(* Logix 5000 project; controller TFF vendor 1 type 14 code 107 rev 33.11; software revision 33.04; part 22 of 38 *)
(* tags used below, declared in another part *)
   Address : DINT;   // Temp Address
   Config : Configuration;   // Index Array used in configuration routines
   Index : DINT;   // Index
   TIME : DINT[2];
   AlarmAnalog : AlarmAnalog[50];   // Analog Alarm Array
   AnalogOutput : AnalogOutput[25];   // Analog Output Array
   AnalogPoint : AnalogInput[50];   // Analog Input Array
   Concentration : Concentration;
   ControlLoop : ControlLoop[20];   // Control Loop Array
   ControlLoop_FeedBagLevel : ALIAS FOR ControlLoop[2];
   ControlLoop_FeedPump : ALIAS FOR ControlLoop[1];
   ControlLoop_TIC101 : ALIAS FOR ControlLoop[7];
   Diafiltration : Diafiltration;
   DigitalPoint : DigitalPoint[150];   // Digital Point Array
   Drive : Drive[11];   // Drives Array
   FQ_Conc : ALIAS FOR Totalizer[0];   // Concentration Totalizer
   FQ_Diaf : ALIAS FOR Totalizer[1];   // DiafiltrationTotalizer
   Mixer : Mixer;   // Mixer config. structure
   Options : Options;   // Options List
   PCV101 : ALIAS FOR AnalogPoint[3];
   Phase : Phases[6];   // Phase Control Array
   Phase0_Totalizer_Feed : ALIAS FOR PhaseTotalizer[0];   // Phase 0 Total Feed
   Phase0_Totalizer_Filtrate : ALIAS FOR PhaseTotalizer[6];   // Phase 0 Total Filtrate
   Phase0_Totalizer_Transfer : ALIAS FOR PhaseTotalizer[12];   // Phase 0 Total Transfer
   Phase1_Totalizer_Feed : ALIAS FOR PhaseTotalizer[1];   // Phase 1 Total Feed
   Phase1_Totalizer_Filtrate : ALIAS FOR PhaseTotalizer[7];   // Phase 1 Total Filtrate
   Phase1_Totalizer_Transfer : ALIAS FOR PhaseTotalizer[13];   // Phase 1 Total Transfer
   Phase2_Totalizer_Feed : ALIAS FOR PhaseTotalizer[2];   // Phase 2 Total Feed
   Phase2_Totalizer_Filtrate : ALIAS FOR PhaseTotalizer[8];   // Phase 2 Total Filtrate
   Phase2_Totalizer_Transfer : ALIAS FOR PhaseTotalizer[14];   // Phase 2 Total Transfer
   Phase3_Totalizer_Feed : ALIAS FOR PhaseTotalizer[3];   // Phase 3 Total Feed
   Phase3_Totalizer_Filtrate : ALIAS FOR PhaseTotalizer[9];   // Phase 3 Total Filtrate
   Phase3_Totalizer_Transfer : ALIAS FOR PhaseTotalizer[15];   // Phase 3 Total Transfer
   Phase4_Totalizer_Feed : ALIAS FOR PhaseTotalizer[4];   // Phase 4 Total Feed
   Phase4_Totalizer_Filtrate : ALIAS FOR PhaseTotalizer[10];   // Phase 4 Total Filtrate
   Phase4_Totalizer_Transfer : ALIAS FOR PhaseTotalizer[16];   // Phase 4 Total Transfer
   Phase5_Totalizer_Feed : ALIAS FOR PhaseTotalizer[5];   // Phase 5 Total Feed
   Phase5_Totalizer_Filtrate : ALIAS FOR PhaseTotalizer[11];   // Phase 5 Total Filtrate
   Phase5_Totalizer_Transfer : ALIAS FOR PhaseTotalizer[17];   // Phase 5 Total Transfer
   Rack_Murr_Node0_Smart : IO_Station;   // Status of Node 0 Smart
   Rack_Murr_Node1_TFF : IO_Station;   // Node 1 data for MOM Config
   Rack_Murr_Node1_TFF20 : IO_Station;   // Status of Node 1 TFF20
   Rack_Murr_Node1_TFF40 : IO_Station;   // Status of Node 1 TFF40
   Rack_Murr_Node1_TFF80 : IO_Station;   // Status of Node 1 TFF80
   SIC002 : ALIAS FOR Drive[2];
   SysControl : SysControl;   // General system status and command
   Tank : TankManagement;   // Tank Management
   ThisSystem : SystemType;
   Valve : Valve[100];   // Valve Array
   ValveControl : ValveControl;   // Valve Control
   XV001 : ALIAS FOR Valve[0];
   XV002 : ALIAS FOR Valve[1];
   XV003 : ALIAS FOR Valve[2];
   XV004 : ALIAS FOR Valve[3];
   XV005 : ALIAS FOR Valve[4];
   XV006 : ALIAS FOR Valve[5];
   XV007 : ALIAS FOR Valve[6];
   XV101 : ALIAS FOR Valve[7];
   XV102 : ALIAS FOR Valve[8];
   XV201 : ALIAS FOR Valve[15];
   XV202 : ALIAS FOR Valve[16];
   XV401 : ALIAS FOR Valve[9];
   XV402 : ALIAS FOR Valve[10];
   XV403 : ALIAS FOR Valve[11];
   XV404 : ALIAS FOR Valve[12];
   XV405 : ALIAS FOR Valve[13];
   XV406 : ALIAS FOR Valve[14];
   XV701 : ALIAS FOR Valve[17];
   XV702 : ALIAS FOR Valve[18];
   XV703 : ALIAS FOR Valve[19];
   XV704 : ALIAS FOR Valve[20];
(* Process, continued *)

ROUTINE Config_IO_Station   (* structured text *)
   (* ==========================================================
   	Config I/O Station : Configure Hardware I/O Cards
   
   	Use 6 output byte for options management.
   		bit 0 to 31 : Enable / Disable 0 to 31 cards (bit index is the module number) --> 0 = Disable
   		bit 32 : Save the configuration --> 1 = Save
   		Buse Control bit 4 : 1 = Switch Off Voltage on modules , 0 = Restart the modules
   
   	List of treatments
   		- Options or configuration tools management
   		- Enable / Disable I/O modules
   		- Switch Off or restart Bus Node
   		- Module Option Management Status
   		- Module Option Management Configuration
   
   -----------------------------------------------------------------------------------------------------------------------------------------------------
   	History
   		2019-DEC-24 - Merck - Q. Spindler - Initial version for Candidate Release 1.00.00.00.a
   ============================================================*)
   
   (*Options or configuration tools management
   ============================================================*)
   
   (* Node 0 *)
   If NOT Rack_Murr_Node0_Smart.MOM_Enable_Config then
   
   	If Options.External_IO then
   		Rack_Murr_Node0_Smart.MOM_Mod_Config[3] := 0 ;
   		Rack_Murr_Node0_Smart.MOM_Mod_Config[4] := 0 ;
   		Rack_Murr_Node0_Smart.MOM_Mod_Config[5] := 0 ;
   		Rack_Murr_Node0_Smart.MOM_Mod_Config[6] := 0 ;
   	else
   		Rack_Murr_Node0_Smart.MOM_Mod_Config[3] := 1 ;
   		Rack_Murr_Node0_Smart.MOM_Mod_Config[4] := 1 ;
   		Rack_Murr_Node0_Smart.MOM_Mod_Config[5] := 1 ;
   		Rack_Murr_Node0_Smart.MOM_Mod_Config[6] := 1 ;
   	End_if ;
   
   		Rack_Murr_Node0_Smart.MOM_Mod_Config[0] := 0 ;
   		Rack_Murr_Node0_Smart.MOM_Mod_Config[1] := 0 ;
   		Rack_Murr_Node0_Smart.MOM_Mod_Config[2] := 0 ;
   		Rack_Murr_Node0_Smart.MOM_Mod_Config[7] := 0 ;
   		Rack_Murr_Node0_Smart.MOM_Mod_Config[8] := 0 ;
   		Rack_Murr_Node0_Smart.MOM_Mod_Config[9] := 0 ;
   		Rack_Murr_Node0_Smart.MOM_Mod_Config[10] := 0 ;
   		Rack_Murr_Node0_Smart.MOM_Mod_Config[11] := 0 ;
   		Rack_Murr_Node0_Smart.MOM_Mod_Config[12] := 0 ;
   		Rack_Murr_Node0_Smart.MOM_Mod_Config[13] := 0 ;
   
   	If Options.FeedTank then
   		Rack_Murr_Node0_Smart.MOM_Mod_Config[14] := 0 ;
   		Rack_Murr_Node0_Smart.MOM_Mod_Config[15] := 0 ;
   		Rack_Murr_Node0_Smart.MOM_Mod_Config[16] := 0 ;
   		Rack_Murr_Node0_Smart.MOM_Mod_Config[17] := 0 ;
   	else
   		Rack_Murr_Node0_Smart.MOM_Mod_Config[14] := 1 ;
   		Rack_Murr_Node0_Smart.MOM_Mod_Config[15] := 1 ;
   		Rack_Murr_Node0_Smart.MOM_Mod_Config[16] := 1 ;
   		Rack_Murr_Node0_Smart.MOM_Mod_Config[17] := 1 ;
   	End_if ;
   		Rack_Murr_Node0_Smart.MOM_Mod_Config[18] := 0 ;
   		Rack_Murr_Node0_Smart.MOM_Mod_Config[19] := 0 ;
   		Rack_Murr_Node0_Smart.MOM_Mod_Config[20] := 0 ;
   		Rack_Murr_Node0_Smart.MOM_Mod_Config[21] := 0 ;
   		Rack_Murr_Node0_Smart.MOM_Mod_Config[22] := 0 ;
   		Rack_Murr_Node0_Smart.MOM_Mod_Config[23] := 0 ;
   		Rack_Murr_Node0_Smart.MOM_Mod_Config[24] := 0 ;
   		Rack_Murr_Node0_Smart.MOM_Mod_Config[25] := 0 ;
   		Rack_Murr_Node0_Smart.MOM_Mod_Config[26] := 0 ;
   		Rack_Murr_Node0_Smart.MOM_Mod_Config[27] := 0 ;
   		Rack_Murr_Node0_Smart.MOM_Mod_Config[28] := 0 ;
   		Rack_Murr_Node0_Smart.MOM_Mod_Config[29] := 0 ;
   		Rack_Murr_Node0_Smart.MOM_Mod_Config[30] := 0 ;
   		Rack_Murr_Node0_Smart.MOM_Mod_Config[31] := 0 ;
   
   End_if ;
   
   
   (* Node 1 *)
   If NOT Rack_Murr_Node1_TFF.MOM_Enable_Config then
   
   	If ThisSystem.MoldType = 123 then
   		Rack_Murr_Node1_TFF.MOM_Mod_Config[0] := 0 ;
   		Rack_Murr_Node1_TFF.MOM_Mod_Config[1] := 0 ;
   		Rack_Murr_Node1_TFF.MOM_Mod_Config[2] := 0 ;
   		Rack_Murr_Node1_TFF.MOM_Mod_Config[3] := 0 ;
   		Rack_Murr_Node1_TFF.MOM_Mod_Config[4] := 0 ;
   		Rack_Murr_Node1_TFF.MOM_Mod_Config[5] := 0 ;
   		Rack_Murr_Node1_TFF.MOM_Mod_Config[6] := 0 ;
   		Rack_Murr_Node1_TFF.MOM_Mod_Config[7] := 0 ;
   		Rack_Murr_Node1_TFF.MOM_Mod_Config[8] := 0 ;
   		Rack_Murr_Node1_TFF.MOM_Mod_Config[9] := 0 ;
   		Rack_Murr_Node1_TFF.MOM_Mod_Config[10] := 0 ;
   		Rack_Murr_Node1_TFF.MOM_Mod_Config[11] := 0 ;
   		Rack_Murr_Node1_TFF.MOM_Mod_Config[12] := 0 ;
   		Rack_Murr_Node1_TFF.MOM_Mod_Config[13] := 0 ;
   		Rack_Murr_Node1_TFF.MOM_Mod_Config[14] := 0 ;
   		Rack_Murr_Node1_TFF.MOM_Mod_Config[15] := 0 ;
   		Rack_Murr_Node1_TFF.MOM_Mod_Config[16] := 0 ;
   		Rack_Murr_Node1_TFF.MOM_Mod_Config[17] := 0 ;
   		Rack_Murr_Node1_TFF.MOM_Mod_Config[18] := 0 ;
   		Rack_Murr_Node1_TFF.MOM_Mod_Config[19] := 0 ;
   		Rack_Murr_Node1_TFF.MOM_Mod_Config[20] := 0 ;
   		Rack_Murr_Node1_TFF.MOM_Mod_Config[21] := 0 ;
   		Rack_Murr_Node1_TFF.MOM_Mod_Config[22] := 0 ;
   		Rack_Murr_Node1_TFF.MOM_Mod_Config[23] := 0 ;
   		Rack_Murr_Node1_TFF.MOM_Mod_Config[24] := 0 ;
   		Rack_Murr_Node1_TFF.MOM_Mod_Config[25] := 0 ;
   		Rack_Murr_Node1_TFF.MOM_Mod_Config[26] := 0 ;
   		Rack_Murr_Node1_TFF.MOM_Mod_Config[27] := 0 ;
   		Rack_Murr_Node1_TFF.MOM_Mod_Config[28] := 0 ;
   		Rack_Murr_Node1_TFF.MOM_Mod_Config[29] := 0 ;
   		Rack_Murr_Node1_TFF.MOM_Mod_Config[30] := 0 ;
   		Rack_Murr_Node1_TFF.MOM_Mod_Config[31] := 0 ;
   	Elsif ThisSystem.MoldType = 124 then
   		Rack_Murr_Node1_TFF.MOM_Mod_Config[0] := 0 ;
   		Rack_Murr_Node1_TFF.MOM_Mod_Config[1] := 0 ;
   		Rack_Murr_Node1_TFF.MOM_Mod_Config[2] := 0 ;
   		Rack_Murr_Node1_TFF.MOM_Mod_Config[3] := 0 ;
   		Rack_Murr_Node1_TFF.MOM_Mod_Config[4] := 0 ;
   		Rack_Murr_Node1_TFF.MOM_Mod_Config[5] := 0 ;
   		Rack_Murr_Node1_TFF.MOM_Mod_Config[6] := 0 ;
   		Rack_Murr_Node1_TFF.MOM_Mod_Config[7] := 0 ;
   		Rack_Murr_Node1_TFF.MOM_Mod_Config[8] := 0 ;
   		Rack_Murr_Node1_TFF.MOM_Mod_Config[9] := 0 ;
   		Rack_Murr_Node1_TFF.MOM_Mod_Config[10] := 0 ;
   		Rack_Murr_Node1_TFF.MOM_Mod_Config[11] := 0 ;
   		Rack_Murr_Node1_TFF.MOM_Mod_Config[12] := 0 ;
   		Rack_Murr_Node1_TFF.MOM_Mod_Config[13] := 0 ;
   		Rack_Murr_Node1_TFF.MOM_Mod_Config[14] := 0 ;
   		Rack_Murr_Node1_TFF.MOM_Mod_Config[15] := 0 ;
   		Rack_Murr_Node1_TFF.MOM_Mod_Config[16] := 0 ;
   		Rack_Murr_Node1_TFF.MOM_Mod_Config[17] := 0 ;
   		Rack_Murr_Node1_TFF.MOM_Mod_Config[18] := 0 ;
   		Rack_Murr_Node1_TFF.MOM_Mod_Config[19] := 0 ;
   		Rack_Murr_Node1_TFF.MOM_Mod_Config[20] := 0 ;
   		Rack_Murr_Node1_TFF.MOM_Mod_Config[21] := 0 ;
   		Rack_Murr_Node1_TFF.MOM_Mod_Config[22] := 0 ;
   		Rack_Murr_Node1_TFF.MOM_Mod_Config[23] := 0 ;
   		Rack_Murr_Node1_TFF.MOM_Mod_Config[24] := 0 ;
   		Rack_Murr_Node1_TFF.MOM_Mod_Config[25] := 0 ;
   		Rack_Murr_Node1_TFF.MOM_Mod_Config[26] := 0 ;
   		Rack_Murr_Node1_TFF.MOM_Mod_Config[27] := 0 ;
   		Rack_Murr_Node1_TFF.MOM_Mod_Config[28] := 0 ;
   		Rack_Murr_Node1_TFF.MOM_Mod_Config[29] := 0 ;
   		Rack_Murr_Node1_TFF.MOM_Mod_Config[30] := 0 ;
   		Rack_Murr_Node1_TFF.MOM_Mod_Config[31] := 0 ;
   	Elsif ThisSystem.MoldType = 126 then
   		Rack_Murr_Node1_TFF.MOM_Mod_Config[0] := 0 ;
   		Rack_Murr_Node1_TFF.MOM_Mod_Config[1] := 0 ;
   		Rack_Murr_Node1_TFF.MOM_Mod_Config[2] := 0 ;
   		Rack_Murr_Node1_TFF.MOM_Mod_Config[3] := 0 ;
   		Rack_Murr_Node1_TFF.MOM_Mod_Config[4] := 0 ;
   		Rack_Murr_Node1_TFF.MOM_Mod_Config[5] := 0 ;
   		Rack_Murr_Node1_TFF.MOM_Mod_Config[6] := 0 ;
   		Rack_Murr_Node1_TFF.MOM_Mod_Config[7] := 0 ;
   		Rack_Murr_Node1_TFF.MOM_Mod_Config[8] := 0 ;
   		Rack_Murr_Node1_TFF.MOM_Mod_Config[9] := 0 ;
   		Rack_Murr_Node1_TFF.MOM_Mod_Config[10] := 0 ;
   		Rack_Murr_Node1_TFF.MOM_Mod_Config[11] := 0 ;
   		Rack_Murr_Node1_TFF.MOM_Mod_Config[12] := 0 ;
   		Rack_Murr_Node1_TFF.MOM_Mod_Config[13] := 0 ;
   		Rack_Murr_Node1_TFF.MOM_Mod_Config[14] := 0 ;
   		Rack_Murr_Node1_TFF.MOM_Mod_Config[15] := 0 ;
   		Rack_Murr_Node1_TFF.MOM_Mod_Config[16] := 0 ;
   		Rack_Murr_Node1_TFF.MOM_Mod_Config[17] := 0 ;
   		Rack_Murr_Node1_TFF.MOM_Mod_Config[18] := 0 ;
   		Rack_Murr_Node1_TFF.MOM_Mod_Config[19] := 0 ;
   		Rack_Murr_Node1_TFF.MOM_Mod_Config[20] := 0 ;
   		Rack_Murr_Node1_TFF.MOM_Mod_Config[21] := 0 ;
   		Rack_Murr_Node1_TFF.MOM_Mod_Config[22] := 0 ;
   		Rack_Murr_Node1_TFF.MOM_Mod_Config[23] := 0 ;
   		Rack_Murr_Node1_TFF.MOM_Mod_Config[24] := 0 ;
   		Rack_Murr_Node1_TFF.MOM_Mod_Config[25] := 0 ;
   		Rack_Murr_Node1_TFF.MOM_Mod_Config[26] := 0 ;
   		Rack_Murr_Node1_TFF.MOM_Mod_Config[27] := 0 ;
   		Rack_Murr_Node1_TFF.MOM_Mod_Config[28] := 0 ;
   		Rack_Murr_Node1_TFF.MOM_Mod_Config[29] := 0 ;
   		Rack_Murr_Node1_TFF.MOM_Mod_Config[30] := 0 ;
   		Rack_Murr_Node1_TFF.MOM_Mod_Config[31] := 0 ;
   	End_if ;
   End_if ;
   
   (*Enable / Disable I/O modules
   ============================================================*)
   
   (* Node 0 *)
   FOR Config.IndexIOMod := 0 to 7 by 1 do
   	RACK_MURR_NODE0_SMART:O.Data[0].[Config.IndexIOMod] := Rack_Murr_Node0_Smart.MOM_Mod_Config[Config.IndexIOMod] ;
   	RACK_MURR_NODE0_SMART:O.Data[1].[Config.IndexIOMod] := Rack_Murr_Node0_Smart.MOM_Mod_Config[Config.IndexIOMod+8] ;
   	RACK_MURR_NODE0_SMART:O.Data[2].[Config.IndexIOMod] := Rack_Murr_Node0_Smart.MOM_Mod_Config[Config.IndexIOMod+16] ;
   	RACK_MURR_NODE0_SMART:O.Data[3].[Config.IndexIOMod] := Rack_Murr_Node0_Smart.MOM_Mod_Config[Config.IndexIOMod+24] ;
   End_for ;
   
   (* Node 1 *)
   FOR Config.IndexIOMod := 0 to 7 by 1 do
   
   	If ThisSystem.MoldType = 123 then
   		RACK_MURR_NODE1_TFF20:O.Data[0].[Config.IndexIOMod] := Rack_Murr_Node1_TFF.MOM_Mod_Config[Config.IndexIOMod] ;
   		RACK_MURR_NODE1_TFF20:O.Data[1].[Config.IndexIOMod] := Rack_Murr_Node1_TFF.MOM_Mod_Config[Config.IndexIOMod+8] ;
   		RACK_MURR_NODE1_TFF20:O.Data[2].[Config.IndexIOMod] := Rack_Murr_Node1_TFF.MOM_Mod_Config[Config.IndexIOMod+16] ;
   		RACK_MURR_NODE1_TFF20:O.Data[3].[Config.IndexIOMod] := Rack_Murr_Node1_TFF.MOM_Mod_Config[Config.IndexIOMod+24] ;
   	Elsif ThisSystem.MoldType = 124 then
   		RACK_MURR_NODE1_TFF40:O.Data[0].[Config.IndexIOMod] := Rack_Murr_Node1_TFF.MOM_Mod_Config[Config.IndexIOMod] ;
   		RACK_MURR_NODE1_TFF40:O.Data[1].[Config.IndexIOMod] := Rack_Murr_Node1_TFF.MOM_Mod_Config[Config.IndexIOMod+8] ;
   		RACK_MURR_NODE1_TFF40:O.Data[2].[Config.IndexIOMod] := Rack_Murr_Node1_TFF.MOM_Mod_Config[Config.IndexIOMod+16] ;
   		RACK_MURR_NODE1_TFF40:O.Data[3].[Config.IndexIOMod] := Rack_Murr_Node1_TFF.MOM_Mod_Config[Config.IndexIOMod+24] ;
   	Elsif ThisSystem.MoldType = 126 then
   		RACK_MURR_NODE1_TFF80:O.Data[0].[Config.IndexIOMod] := Rack_Murr_Node1_TFF.MOM_Mod_Config[Config.IndexIOMod] ;
   		RACK_MURR_NODE1_TFF80:O.Data[1].[Config.IndexIOMod] := Rack_Murr_Node1_TFF.MOM_Mod_Config[Config.IndexIOMod+8] ;
   		RACK_MURR_NODE1_TFF80:O.Data[2].[Config.IndexIOMod] := Rack_Murr_Node1_TFF.MOM_Mod_Config[Config.IndexIOMod+16] ;
   		RACK_MURR_NODE1_TFF80:O.Data[3].[Config.IndexIOMod] := Rack_Murr_Node1_TFF.MOM_Mod_Config[Config.IndexIOMod+24] ;
   	End_if ;
   
   End_for ;
   
   (* Switch Off or restart Bus Node
   ============================================================*)
   
   (* Node 0 *)
   RACK_MURR_NODE0_SMART:O.Data[6].4 := Rack_Murr_Node0_Smart.MOM_Restart ;
   
   (* Node 1 *)
   If ThisSystem.MoldType = 123 then
   	RACK_MURR_NODE1_TFF20:O.Data[6].4 := Rack_Murr_Node1_TFF.MOM_Restart ;
   Elsif ThisSystem.MoldType = 124 then
   	RACK_MURR_NODE1_TFF40:O.Data[6].4 := Rack_Murr_Node1_TFF.MOM_Restart ;
   Elsif ThisSystem.MoldType = 126 then
   	RACK_MURR_NODE1_TFF80:O.Data[6].4 := Rack_Murr_Node1_TFF.MOM_Restart ;
   End_if ;
   
   (* Module Option Management Status
   ============================================================*)
   (* Node 0 *)
   Rack_Murr_Node0_Smart.MOM_Status := RACK_MURR_NODE0_SMART:I.Data[0];
   
   (* Node 1 *)
   If ThisSystem.MoldType = 123 then
   	Rack_Murr_Node1_TFF.MOM_Status := RACK_MURR_NODE1_TFF20:I.Data[0];
   Elsif ThisSystem.MoldType = 124 then
   	Rack_Murr_Node1_TFF.MOM_Status := RACK_MURR_NODE1_TFF40:I.Data[0];
   Elsif ThisSystem.MoldType = 126 then
   	Rack_Murr_Node1_TFF.MOM_Status := RACK_MURR_NODE1_TFF80:I.Data[0];
   End_if ;
   
   (*Module Option Management Configuration
   ============================================================*)
   
   (*save the Module Option Management configuration*)
   
   (* Node 0 *)
   RACK_MURR_NODE0_SMART:O.Data[4].0 := 1 ;
   
   (* Node 1 *)
   If ThisSystem.MoldType = 123 then
   	RACK_MURR_NODE1_TFF20:O.Data[4].0 := 1 ;
   Elsif ThisSystem.MoldType = 124 then
   	RACK_MURR_NODE1_TFF40:O.Data[4].0 := 1 ;
   Elsif ThisSystem.MoldType = 126 then
   	RACK_MURR_NODE1_TFF80:O.Data[4].0 := 1 ;
   End_if ;
   
END_ROUTINE

ROUTINE Config_Options   (* structured text *)
   (* ==========================================================
   	Config Options : Configure Options
   
   	List of treatments
   		- Configure Automatic options
   		- Configure Tank options
   		- Configure Flag for current installed clamshell
   
   -----------------------------------------------------------------------------------------------------------------------------------------------------
   	History
   		2019-DEC-24 - Merck - Q. Spindler - Initial version for Candidate Release 1.00.00.00.a
   		2022-SEP-22 - Actemium - J. Jaekel - Modification for Candidate Release 1.01.00.01.a
   				- Add Magnetic Filtrate Flowmeter instead of Ultrasonic option
   ============================================================*)
   
   (*Configure options if option Simulation mode is disabled*)
   IF Not SysControl.Simulate_Options THEN
   	// Inlet Feed Disable Option
   	IF Options.InletFeed THEN
   		Options.InletFeed_Dis := 0;
   	ELSE
   		Options.InletFeed_Dis := 1;
   	END_IF;
   
   	// No Instrum Disable Option
   	IF Options.FiltrateNoInstrum THEN
   		Options.FiltrateNoInstrum_Dis := 0;
   	ELSE
   		Options.FiltrateNoInstrum_Dis := 1;
   	END_IF;
   
   	// Tank Option
   	IF NOT Options.FeedTank THEN
   		Options.TankPH := 0;
   		Options.TankCond := 0;
   	END_IF;
   
   	// Single Use Option
   	IF Options.FiltrateNoInstrum THEN
   		Options.SingleUsePH := 0;
   	END_IF;
   
   	// Magnetic Filtrate Flowmeter instead of Ultrasonic
   	IF Options.FiltrateUltrasonicFlow THEN
   		Options.FiltrateMagneticFlow := 0;
   	ELSE
   		Options.FiltrateMagneticFlow := 1;
   	END_IF;
   END_IF;
   
   
   (*Simulate Tank Range*)
   IF Tank.Config.Simulate THEN
   
   	CASE	Tank.Config.Option_Simulate OF
   		0:	Tank.Config.Option_Current := 0 ;
   		1:	Tank.Config.Option_Current := 1 ;
   		2:	Tank.Config.Option_Current := 2 ;
   		3:	Tank.Config.Option_Current := 3 ;
   	ELSE 	Tank.Config.Option_Current := 0 ;
   	END_CASE;
   
   END_IF;
   
   (* Configure Flag for current installed clamshell
   Used to create the CCP Configuration file based on current clamshell
   ============================================================*)
   IF ThisSystem.MoldType = 123 THEN
   
   	Options.TFF20 := 1 ;
   	Options.TFF40 := 0 ;
   	Options.TFF80 := 0 ;
   
   ELSIF ThisSystem.MoldType = 124 THEN
   
   	Options.TFF20 := 0 ;
   	Options.TFF40 := 1 ;
   	Options.TFF80 := 0 ;
   
   ELSIF ThisSystem.MoldType = 126 THEN
   
   	Options.TFF20 := 0 ;
   	Options.TFF40 := 0 ;
   	Options.TFF80 := 1 ;
   
   END_IF;
END_ROUTINE

ROUTINE Config_Reset   (* structured text *)
// Set to 0  all settings
   (* ==========================================================
   	Config Reset : 	When config.reset command is activated,AnalogPoint, AlarmAnalog, AnalogOutput, Drive, DigitalPoint and Valve structure
   					are initialized to 0.
   
   	List of treatments
   		- AnalogPoint Structure reset [0] to [49]
   		- AlarmAnalog Structure reset [0] to [49]
   		- AnalogOutput Structure reset [0] to [24]
   		- Drive Structure reset [0] to [10]
   		- DigitalPoint Structure reset [0] to [149]
   		- Valve Structure reset [0] to [99]
   
   -----------------------------------------------------------------------------------------------------------------------------------------------------
   	History
   		2019-DEC-24 - Merck - Q. Spindler - Initial version for Candidate Release 1.00.00.00.a
   ============================================================*)
   
   
   (*Structure Reset [0] to [149]
   ============================================================*)
   IF Config.Reset THEN
   	FOR Config.IndexReset := 0 TO 149 BY 1 Do
   		IF Config.IndexReset <= 49 THEN
   		(*AnalogPoint Structure Reset [0] to [49]
   		====================================================*)
   			AnalogPoint[Config.IndexReset].OutofRange := 0 ;
   			AnalogPoint[Config.IndexReset].FilterType := 0 ;
   			AnalogPoint[Config.IndexReset].AveragingTotal := 0 ;
   			AnalogPoint[Config.IndexReset].Address := 0 ;
   			AnalogPoint[Config.IndexReset].RawMin := 0 ;
   			AnalogPoint[Config.IndexReset].RawMax := 0 ;
   			AnalogPoint[Config.IndexReset].RawValue := 0 ;
   			AnalogPoint[Config.IndexReset].RawLowLimit := 0 ;
   			AnalogPoint[Config.IndexReset].RawHighLimit := 0 ;
   			AnalogPoint[Config.IndexReset].FilterUser := 0 ;
   			AnalogPoint[Config.IndexReset].FilteredRaw := 0 ;
   			AnalogPoint[Config.IndexReset].FilterActual := 0 ;
   			AnalogPoint[Config.IndexReset].ScaledMin := 0 ;
   			AnalogPoint[Config.IndexReset].ScaledMax := 0 ;
   			AnalogPoint[Config.IndexReset].RangeMin := 0 ;
   			AnalogPoint[Config.IndexReset].RangeMax := 0 ;
   			AnalogPoint[Config.IndexReset].RangeMinSave := 0 ;
   			AnalogPoint[Config.IndexReset].RangeMaxSave := 0 ;
   			AnalogPoint[Config.IndexReset].RealCfg := 0 ;
   			AnalogPoint[Config.IndexReset].EnableCfg := 0 ;
   			AnalogPoint[Config.IndexReset].OverrideCfg := 0 ;
   
   		(*AlarmAnalog Structure Reset [0] to [49]
   		====================================================*)
   			AlarmAnalog[Config.IndexReset].Override := 0 ;
   			AlarmAnalog[Config.IndexReset].Disable := 0 ;
   			AlarmAnalog[Config.IndexReset].LOLODisable := 0 ;
   			AlarmAnalog[Config.IndexReset].LODisable := 0 ;
   			AlarmAnalog[Config.IndexReset].HIDisable := 0 ;
   			AlarmAnalog[Config.IndexReset].HIHIDisable := 0 ;
   			AlarmAnalog[Config.IndexReset].HIHIEnable := 0 ;
   			AlarmAnalog[Config.IndexReset].FeedPumpEnable := 0 ;
   			AlarmAnalog[Config.IndexReset].FeedPumpTag := 0 ;
   			AlarmAnalog[Config.IndexReset].TransferPumpEnable := 0 ;
   			AlarmAnalog[Config.IndexReset].TransferPumpTag := 0 ;
   			AlarmAnalog[Config.IndexReset].LOLO := 0 ;
   			AlarmAnalog[Config.IndexReset].LO := 0 ;
   			AlarmAnalog[Config.IndexReset].HI := 0 ;
   			AlarmAnalog[Config.IndexReset].HIHI := 0 ;
   			AlarmAnalog[Config.IndexReset].LOLOTimer.PRE := 0 ;
   			AlarmAnalog[Config.IndexReset].LOTimer.PRE := 0 ;
   			AlarmAnalog[Config.IndexReset].HITimer.PRE := 0 ;
   			AlarmAnalog[Config.IndexReset].HIHITimer.PRE := 0 ;
   			AlarmAnalog[Config.IndexReset].EnableCfg := 0 ;
   		End_IF;
   
   		(*AnalogOutput Structure Reset [0] to [24]
   		====================================================*)
   		IF Config.IndexReset <= 24 THEN
   			AnalogOutput[Config.IndexReset].RawValue := 0 ;
   			AnalogOutput[Config.IndexReset].RawMin := 0 ;
   			AnalogOutput[Config.IndexReset].RawMax := 0 ;
   			AnalogOutput[Config.IndexReset].ScaledMin := 0 ;
   			AnalogOutput[Config.IndexReset].ScaledMax := 0 ;
   			AnalogOutput[Config.IndexReset].EnableCfg := 0 ;
   		End_IF;
   
   		(*Drive Structure Reset [0] to [10]
   		====================================================*)
   		IF Config.IndexReset <= 10 THEN
   			Drive[Config.IndexReset].OutputAddress := 0 ;
   			Drive[Config.IndexReset].InputAddress := 0 ;
   			Drive[Config.IndexReset].RunInput := 0 ;
   			Drive[Config.IndexReset].InterlockTimer.PRE := 0 ;
   			Drive[Config.IndexReset].EnableCfg := 0 ;
   			Drive[Config.IndexReset].ReverseCfg := 0 ;
   			Drive[Config.IndexReset].Direction := 0 ;
   			Drive[Config.IndexReset].DirectionAddress := 0 ;
   		End_IF;
   
   		IF Config.IndexReset <= 99 THEN
   				(*Valves Structure Reset [0] to [99]
   		====================================================*)
   		Valve[Config.IndexReset].ZSOpenEnable := 0 ;
   		Valve[Config.IndexReset].ZSCloseEnable := 0 ;
   		Valve[Config.IndexReset].ZSOverride := 0 ;
   		Valve[Config.IndexReset].FailState := 0 ;
   		Valve[Config.IndexReset].Ports := 0 ;
   		Valve[Config.IndexReset].EnableCfg := 0 ;
   		Valve[Config.IndexReset].StatusWord := 0 ;
   		Valve[Config.IndexReset].ZSOpenAddress := 0 ;
   		Valve[Config.IndexReset].ZSCloseAddress := 0 ;
   		Valve[Config.IndexReset].OutputAddress := 0 ;
   		Valve[Config.IndexReset].AlarmTimer.PRE := 0 ;
   		Valve[Config.IndexReset].AutoCloseTimer.PRE := 0 ;
   		End_IF;
   
   		(*DigitalPoint Structure Reset [0] to [149]
   		====================================================*)
   		DigitalPoint[Config.IndexReset].Override := 0 ;
   		DigitalPoint[Config.IndexReset].DelayTimer.PRE := 0 ;
   		DigitalPoint[Config.IndexReset].Priority := 0 ;
   		DigitalPoint[Config.IndexReset].EnableCfg := 0 ;
   		DigitalPoint[Config.IndexReset].ActiveStateCFg := 0 ;
   		DigitalPoint[Config.IndexReset].RealInputCfg := 0 ;
   		DigitalPoint[Config.IndexReset].InputAddressCfg := 0 ;
   		DigitalPoint[Config.IndexReset].AlarmCfg := 0 ;
   		DigitalPoint[Config.IndexReset].AlarmStateCfg := 0 ;
   		DigitalPoint[Config.IndexReset].OverrideCfg := 0 ;
   		DigitalPoint[Config.IndexReset].PriorityCfg := 0 ;
   		DigitalPoint[Config.IndexReset].Cond1Cfg := 0 ;
   		DigitalPoint[Config.IndexReset].Cond2Cfg := 0 ;
   		DigitalPoint[Config.IndexReset].FlashingInputCfg := 0 ;
   
   	END_FOR;
   End_IF;
   (*Reset config.reset to execute routine one time*)
   Config.Reset := 0;
END_ROUTINE

ROUTINE Config_Totalizers   (* structured text *)
   (* ==========================================================
   	Config Totalizers : Configure Totalizers Structure
   
   	List of treatments
   		- Phase 0 Totalizers
   		- Phase 1 Totalizers
   		- Phase 2 Totalizers
   		- Phase 3 Totalizers
   		- Phase 4 Totalizers
   		- Phase 5 Totalizers
   		- Concentration and Diafiltration Totalizers
   
   -----------------------------------------------------------------------------------------------------------------------------------------------------
   	History
   		2019-DEC-24 - Merck - Q. Spindler - Initial version for Candidate Release 1.00.00.00.a
   		2022-JAN-11 - Merck - Q. Spindler - Modifications for Candidate Release 1.01.00.00.a
   					- Add transfer totalizers
   ============================================================*)
   
   
   (*Phase 0 Totalizers
   ============================================================*)
   Phase0_Totalizer_Feed.EnableCfg := 1 ;
   Phase0_Totalizer_Feed.SourceAddressCfg := 42 ;
   Phase0_Totalizer_Feed.SourceTypeCfg := 0 ;
   Phase0_Totalizer_Feed.PVscale := 60 ;
   
   Phase0_Totalizer_Filtrate.EnableCfg := 1 ;
   Phase0_Totalizer_Filtrate.SourceAddressCfg := 2 ;
   Phase0_Totalizer_Filtrate.SourceTypeCfg := 0 ;
   Phase0_Totalizer_Filtrate.PVscale := 60 ;
   
   Phase0_Totalizer_Transfer.EnableCfg := 1 ;
   Phase0_Totalizer_Transfer.SourceAddressCfg := 20 ;
   Phase0_Totalizer_Transfer.SourceTypeCfg := 0 ;
   Phase0_Totalizer_Transfer.PVscale := 60 ;
   
   (*Phase 1 Totalizers
   ============================================================*)
   Phase1_Totalizer_Feed.EnableCfg := 1 ;
   Phase1_Totalizer_Feed.SourceAddressCfg := 42 ;
   Phase1_Totalizer_Feed.SourceTypeCfg := 0 ;
   Phase1_Totalizer_Feed.PVscale := 60 ;
   
   Phase1_Totalizer_Filtrate.EnableCfg := 1 ;
   Phase1_Totalizer_Filtrate.SourceAddressCfg := 2 ;
   Phase1_Totalizer_Filtrate.SourceTypeCfg := 0 ;
   Phase1_Totalizer_Filtrate.PVscale := 60 ;
   
   Phase1_Totalizer_Transfer.EnableCfg := 1 ;
   Phase1_Totalizer_Transfer.SourceAddressCfg := 20 ;
   Phase1_Totalizer_Transfer.SourceTypeCfg := 0 ;
   Phase1_Totalizer_Transfer.PVscale := 60 ;
   
   (*Phase 2 Totalizers
   ============================================================*)
   Phase2_Totalizer_Feed.EnableCfg := 1 ;
   Phase2_Totalizer_Feed.SourceAddressCfg := 42 ;
   Phase2_Totalizer_Feed.SourceTypeCfg := 0 ;
   Phase2_Totalizer_Feed.PVscale := 60 ;
   
   Phase2_Totalizer_Filtrate.EnableCfg := 1 ;
   Phase2_Totalizer_Filtrate.SourceAddressCfg := 2 ;
   Phase2_Totalizer_Filtrate.SourceTypeCfg := 0 ;
   Phase2_Totalizer_Filtrate.PVscale := 60 ;
   
   Phase2_Totalizer_Transfer.EnableCfg := 1 ;
   Phase2_Totalizer_Transfer.SourceAddressCfg := 20 ;
   Phase2_Totalizer_Transfer.SourceTypeCfg := 0 ;
   Phase2_Totalizer_Transfer.PVscale := 60 ;
   
   (*Phase 3 Totalizers
   ============================================================*)
   Phase3_Totalizer_Feed.EnableCfg := 1 ;
   Phase3_Totalizer_Feed.SourceAddressCfg := 42 ;
   Phase3_Totalizer_Feed.SourceTypeCfg := 0 ;
   Phase3_Totalizer_Feed.PVscale := 60 ;
   
   Phase3_Totalizer_Filtrate.EnableCfg := 1 ;
   Phase3_Totalizer_Filtrate.SourceAddressCfg := 2 ;
   Phase3_Totalizer_Filtrate.SourceTypeCfg := 0 ;
   Phase3_Totalizer_Filtrate.PVscale := 60 ;
   
   Phase3_Totalizer_Transfer.EnableCfg := 1 ;
   Phase3_Totalizer_Transfer.SourceAddressCfg := 20 ;
   Phase3_Totalizer_Transfer.SourceTypeCfg := 0 ;
   Phase3_Totalizer_Transfer.PVscale := 60 ;
   
   (*Phase 4 Totalizers
   ============================================================*)
   Phase4_Totalizer_Feed.EnableCfg := 1 ;
   Phase4_Totalizer_Feed.SourceAddressCfg := 42 ;
   Phase4_Totalizer_Feed.SourceTypeCfg := 0 ;
   Phase4_Totalizer_Feed.PVscale := 60 ;
   
   Phase4_Totalizer_Filtrate.EnableCfg := 1 ;
   Phase4_Totalizer_Filtrate.SourceAddressCfg := 2 ;
   Phase4_Totalizer_Filtrate.SourceTypeCfg := 0 ;
   Phase4_Totalizer_Filtrate.PVscale := 60 ;
   
   Phase4_Totalizer_Transfer.EnableCfg := 1 ;
   Phase4_Totalizer_Transfer.SourceAddressCfg := 20 ;
   Phase4_Totalizer_Transfer.SourceTypeCfg := 0 ;
   Phase4_Totalizer_Transfer.PVscale := 60 ;
   
   (*Phase 5 Totalizers
   ============================================================*)
   Phase5_Totalizer_Feed.EnableCfg := 1 ;
   Phase5_Totalizer_Feed.SourceAddressCfg := 42 ;
   Phase5_Totalizer_Feed.SourceTypeCfg := 0 ;
   Phase5_Totalizer_Feed.PVscale := 60 ;
   
   Phase5_Totalizer_Filtrate.EnableCfg := 1 ;
   Phase5_Totalizer_Filtrate.SourceAddressCfg := 2 ;
   Phase5_Totalizer_Filtrate.SourceTypeCfg := 0 ;
   Phase5_Totalizer_Filtrate.PVscale := 60 ;
   
   Phase5_Totalizer_Transfer.EnableCfg := 1 ;
   Phase5_Totalizer_Transfer.SourceAddressCfg := 20 ;
   Phase5_Totalizer_Transfer.SourceTypeCfg := 0 ;
   Phase5_Totalizer_Transfer.PVscale := 60 ;
   
   (*Concentration and Diafiltration Totalizers
   ============================================================*)
   
   FQ_Conc.PVscale := 60 ;
   FQ_Diaf.PVscale := 60 ;
END_ROUTINE

ROUTINE Config_Valve   (* structured text *)
// Apply the default configuration
   (* ==========================================================
   	Config Valve : Configure Valve Structure
   
   	List of treatments
   		- Valve[0] : Valve XV001
   		- Valve[1] : Valve XV002
   		- Valve[2] : Valve XV003
   		- Valve[3] : Valve XV004
   		- Valve[4] : Valve XV005
   		- Valve[5] : Valve XV006
   		- Valve[6] : Valve XV007
   		- Valve[7] : Valve XV101
   		- Valve[8] : Valve XV102
   		- Valve[9] : Valve XV401
   		- Valve[10]: Valve XV402
   		- Valve[11]: Valve XV403
   		- Valve[12]: Valve XV404
   		- Valve[13]: Valve XV405
   		- Valve[14]: Valve XV406
   		- Valve[15]: Valve XV201
   		- Valve[16]: Valve XV202
   		- Valve[17]: Valve XV701
   		- Valve[18]: Valve XV702
   		- Valve[19]: Valve XV703
   		- Valve[20]: Valve XV704
   		- Reset Loop : Set to 0 the Valve[21 to 99].EnableCfg
   
   -----------------------------------------------------------------------------------------------------------------------------------------------------
   	History
   		2019-DEC-24 - Merck - Q. Spindler - Initial version for Candidate Release 1.00.00.00.a
   		2020-APR-06 - Merck - Q. Spindler - Modifications for Candidate Release 1.00.00.00.b
   					- Invert FailState for XV201
   					- Add ZSClose for XV003,XV004,XV005,XV006,XV007
   		2020-JUN-19 - Merck - Q. Spindler - Modifications for Candidate Release 1.00.00.00.c
   					- Change ZSClose to ZSOpen for XV003,XV004,XV005,XV006,XV007
   ============================================================*)
   
   
   (*Max valve number use as terminal value in loop
   ============================================================*)
   ValveControl.MaxValveNum := 32;
   
   (*Valve[0] : Valve XV001
   ============================================================*)
   Valve[0].EnableCfg := 1 ;
   Valve[0].FailState := 1 ;
   Valve[0].ZSOverride := 1 ;
   Valve[0].Ports := 0 ;
   Valve[0].PriorityCfg := 0 ;
   Valve[0].ZSOpenEnable := 0 ;
   Valve[0].Alarm := 0 ;
   Valve[0].ZSCloseEnable := 0 ;
   Valve[0].ZSOpenAddress := 0 ;
   Valve[0].ZSCloseAddress := 0 ;
   Valve[0].OutputAddress := 32 ;
   
   (*Valve[1] : Valve XV002
   ============================================================*)
   Valve[1].EnableCfg := 1 ;
   Valve[1].FailState := 1 ;
   Valve[1].ZSOverride := 1 ;
   Valve[1].Ports := 0 ;
   Valve[1].PriorityCfg := 0 ;
   Valve[1].ZSOpenEnable := 0 ;
   Valve[1].Alarm := 0 ;
   Valve[1].ZSCloseEnable := 0 ;
   Valve[1].ZSOpenAddress := 0 ;
   Valve[1].ZSCloseAddress := 0 ;
   Valve[1].OutputAddress := 33 ;
   
   (*Valve[2] : Valve XV003
   ============================================================*)
   IF Options.InletFeed THEN
   	Valve[2].EnableCfg := 1 ;
   ELSE
   	Valve[2].EnableCfg := 0 ;
   	Valve[2].Alarm := 0 ;
   END_IF;
   Valve[2].FailState := 0 ;
   Valve[2].Ports := 0 ;
   Valve[2].PriorityCfg := 1 ;
   Valve[2].ZSOpenEnable := 1 ;
   Valve[2].ZSCloseEnable := 0 ;
   Valve[2].ZSOpenAddress := 2 ;
   Valve[2].ZSCloseAddress := 0 ;
   Valve[2].OutputAddress := 34 ;
   
   (*Valve[3] : Valve XV004
   ============================================================*)
   IF Options.InletFeed THEN
   	Valve[3].EnableCfg := 1 ;
   ELSE
   	Valve[3].EnableCfg := 0 ;
   	Valve[3].Alarm := 0 ;
   END_IF;
   Valve[3].FailState := 0 ;
   Valve[3].Ports := 0 ;
   Valve[3].PriorityCfg := 1 ;
   Valve[3].ZSOpenEnable := 1 ;
   Valve[3].ZSCloseEnable := 0 ;
   Valve[3].ZSOpenAddress := 3 ;
   Valve[3].ZSCloseAddress := 0 ;
   Valve[3].OutputAddress := 35 ;
   
   (*Valve[4] : Valve XV005
   ============================================================*)
   IF Options.InletFeed THEN
   	Valve[4].EnableCfg := 1 ;
   ELSE
   	Valve[4].EnableCfg := 0 ;
   	Valve[4].Alarm := 0 ;
   END_IF;
   Valve[4].FailState := 0 ;
   Valve[4].Ports := 0 ;
   Valve[4].PriorityCfg := 1 ;
   Valve[4].ZSOpenEnable := 1 ;
   Valve[4].ZSCloseEnable := 0 ;
   Valve[4].ZSOpenAddress := 4 ;
   Valve[4].ZSCloseAddress := 0 ;
   Valve[4].OutputAddress := 36 ;
   
   (*Valve[5] : Valve XV006
   ============================================================*)
   IF Options.InletFeed THEN
   	Valve[5].EnableCfg := 1 ;
   ELSE
   	Valve[5].EnableCfg := 0 ;
   	Valve[5].Alarm := 0 ;
   END_IF;
   Valve[5].FailState := 0 ;
   Valve[5].Ports := 0 ;
   Valve[5].PriorityCfg := 1 ;
   Valve[5].ZSOpenEnable := 1 ;
   Valve[5].ZSCloseEnable := 0 ;
   Valve[5].ZSOpenAddress := 5 ;
   Valve[5].ZSCloseAddress := 0 ;
   Valve[5].OutputAddress := 37 ;
   
   (*Valve[6] : Valve XV007
   ============================================================*)
   IF Options.InletFeed THEN
   	Valve[6].EnableCfg := 1 ;
   ELSE
   	Valve[6].EnableCfg := 0 ;
   	Valve[6].Alarm := 0 ;
   END_IF;
   Valve[6].FailState := 0 ;
   Valve[6].Ports := 0 ;
   Valve[6].PriorityCfg := 1 ;
   Valve[6].ZSOpenEnable := 1 ;
   Valve[6].ZSCloseEnable := 0 ;
   Valve[6].ZSOpenAddress := 6;
   Valve[6].ZSCloseAddress := 0 ;
   Valve[6].OutputAddress := 38 ;
   
   (*Valve[7] : Valve XV101
   ============================================================*)
   Valve[7].EnableCfg := 1 ;
   Valve[7].FailState := 1 ;
   Valve[7].ZSOverride := 1 ;
   Valve[7].Ports := 0 ;
   Valve[7].PriorityCfg := 0 ;
   Valve[7].ZSOpenEnable := 0 ;
   Valve[7].Alarm := 0 ;
   Valve[7].ZSCloseEnable := 0 ;
   Valve[7].ZSOpenAddress := 0 ;
   Valve[7].ZSCloseAddress := 0 ;
   Valve[7].OutputAddress := 39 ;
   
   (*Valve[8] : Valve XV102
   ============================================================*)
   Valve[8].EnableCfg := 1 ;
   Valve[8].FailState := 1 ;
   Valve[8].ZSOverride := 1 ;
   Valve[8].Ports := 0 ;
   Valve[8].PriorityCfg := 0 ;
   Valve[8].ZSOpenEnable := 0 ;
   Valve[8].Alarm := 0 ;
   Valve[8].ZSCloseEnable := 0 ;
   Valve[8].ZSOpenAddress := 0 ;
   Valve[8].ZSCloseAddress := 0 ;
   Valve[8].OutputAddress := 40 ;
   
   (*Valve[9] : Valve XV401
   ============================================================*)
   Valve[9].EnableCfg := 1 ;
   Valve[9].FailState := 0 ;
   Valve[9].ZSOverride := 1 ;
   Valve[9].Ports := 0 ;
   Valve[9].PriorityCfg := 0 ;
   Valve[9].ZSOpenEnable := 0 ;
   Valve[9].Alarm := 0 ;
   Valve[9].ZSCloseEnable := 0 ;
   Valve[9].ZSOpenAddress := 0 ;
   Valve[9].ZSCloseAddress := 0 ;
   Valve[9].OutputAddress := 41 ;
   
   (*Valve[10]: Valve XV402
   ============================================================*)
   Valve[10].EnableCfg := 1 ;
   Valve[10].FailState := 0 ;
   Valve[10].ZSOverride := 1 ;
   Valve[10].Ports := 0 ;
   Valve[10].PriorityCfg := 0 ;
   Valve[10].ZSOpenEnable := 0 ;
   Valve[10].Alarm := 0 ;
   Valve[10].ZSCloseEnable := 0 ;
   Valve[10].ZSOpenAddress := 0 ;
   Valve[10].ZSCloseAddress := 0 ;
   Valve[10].OutputAddress := 42 ;
   
   (*Valve[11]: Valve XV403
   ============================================================*)
   Valve[11].EnableCfg := 1 ;
   Valve[11].FailState := 0 ;
   Valve[11].ZSOverride := 1 ;
   Valve[11].Ports := 0 ;
   Valve[11].PriorityCfg := 0 ;
   Valve[11].ZSOpenEnable := 0 ;
   Valve[11].Alarm := 0 ;
   Valve[11].ZSCloseEnable := 0 ;
   Valve[11].ZSOpenAddress := 0 ;
   Valve[11].ZSCloseAddress := 0 ;
   Valve[11].OutputAddress := 43 ;
   
   (*Valve[12]: Valve XV404
   ============================================================*)
   Valve[12].EnableCfg := 1 ;
   Valve[12].FailState := 0 ;
   Valve[12].ZSOverride := 1 ;
   Valve[12].Ports := 0 ;
   Valve[12].PriorityCfg := 0 ;
   Valve[12].ZSOpenEnable := 0 ;
   Valve[12].Alarm := 0 ;
   Valve[12].ZSCloseEnable := 0 ;
   Valve[12].ZSOpenAddress := 0 ;
   Valve[12].ZSCloseAddress := 0 ;
   Valve[12].OutputAddress := 44 ;
   
   (*Valve[13]: Valve XV405
   ============================================================*)
   IF Options.InletFeed THEN
   	Valve[13].EnableCfg := 0 ;
   ELSE
   	Valve[13].EnableCfg := 1 ;
   END_IF;
   Valve[13].FailState := 0 ;
   Valve[13].ZSOverride := 1 ;
   Valve[13].Ports := 0 ;
   Valve[13].PriorityCfg := 0 ;
   Valve[13].ZSOpenEnable := 0 ;
   Valve[13].Alarm := 0 ;
   Valve[13].ZSCloseEnable := 0 ;
   Valve[13].ZSOpenAddress := 0 ;
   Valve[13].ZSCloseAddress := 0 ;
   Valve[13].OutputAddress := 45 ;
   
   (*Valve[14]: Valve XV406
   ============================================================*)
   IF Options.InletFeed THEN
   	Valve[14].EnableCfg := 0 ;
   ELSE
   	Valve[14].EnableCfg := 1 ;
   END_IF;
   Valve[14].FailState := 0 ;
   Valve[14].ZSOverride := 1 ;
   Valve[14].Ports := 0 ;
   Valve[14].PriorityCfg := 0 ;
   Valve[14].ZSOpenEnable := 0 ;
   Valve[14].Alarm := 0 ;
   Valve[14].ZSCloseEnable := 0 ;
   Valve[14].ZSOpenAddress := 0 ;
   Valve[14].ZSCloseAddress := 0 ;
   Valve[14].OutputAddress := 46 ;
   
   (*Valve[15]: Valve XV201
   ============================================================*)
   Valve[15].EnableCfg := 1 ;
   Valve[15].FailState := 0 ;
   Valve[15].ZSOverride := 1 ;
   Valve[15].Ports := 0 ;
   Valve[15].PriorityCfg := 0 ;
   Valve[15].ZSOpenEnable := 0 ;
   Valve[15].Alarm := 0 ;
   Valve[15].ZSCloseEnable := 0 ;
   Valve[15].ZSOpenAddress := 0 ;
   Valve[15].ZSCloseAddress := 0 ;
   Valve[15].OutputAddress := 47 ;
   
   (*Valve[16]: Valve XV202
   ============================================================*)
   Valve[16].EnableCfg := 1 ;
   Valve[16].FailState := 0 ;
   Valve[16].ZSOverride := 1 ;
   Valve[16].Ports := 0 ;
   Valve[16].PriorityCfg := 0 ;
   Valve[16].ZSOpenEnable := 0 ;
   Valve[16].Alarm := 0 ;
   Valve[16].ZSCloseEnable := 0 ;
   Valve[16].ZSOpenAddress := 0 ;
   Valve[16].ZSCloseAddress := 0 ;
   Valve[16].OutputAddress := 48 ;
   
   (*Valve[17]: Valve XV701
   ============================================================*)
   Valve[17].EnableCfg := 1 ;
   Valve[17].FailState := 0 ;
   Valve[17].ZSOverride := 1 ;
   Valve[17].Ports := 0 ;
   Valve[17].PriorityCfg := 0 ;
   Valve[17].ZSOpenEnable := 0 ;
   Valve[17].Alarm := 0 ;
   Valve[17].ZSCloseEnable := 0 ;
   Valve[17].ZSOpenAddress := 0 ;
   Valve[17].ZSCloseAddress := 0 ;
   Valve[17].OutputAddress := 49 ;
   
   (*Valve[18]: Valve XV702
   ============================================================*)
   Valve[18].EnableCfg := 1 ;
   Valve[18].FailState := 0 ;
   Valve[18].ZSOverride := 1 ;
   Valve[18].Ports := 0 ;
   Valve[18].PriorityCfg := 0 ;
   Valve[18].ZSOpenEnable := 0 ;
   Valve[18].Alarm := 0 ;
   Valve[18].ZSCloseEnable := 0 ;
   Valve[18].ZSOpenAddress := 0 ;
   Valve[18].ZSCloseAddress := 0 ;
   Valve[18].OutputAddress := 50 ;
   
   (*Valve[19]: Valve XV703
   ============================================================*)
   Valve[19].EnableCfg := 1 ;
   Valve[19].FailState := 0 ;
   Valve[19].ZSOverride := 1 ;
   Valve[19].Ports := 0 ;
   Valve[19].PriorityCfg := 0 ;
   Valve[19].ZSOpenEnable := 0 ;
   Valve[19].Alarm := 0 ;
   Valve[19].ZSCloseEnable := 0 ;
   Valve[19].ZSOpenAddress := 0 ;
   Valve[19].ZSCloseAddress := 0 ;
   Valve[19].OutputAddress := 51 ;
   
   (*Valve[20]: Valve XV704
   ============================================================*)
   Valve[20].EnableCfg := 1 ;
   Valve[20].FailState := 0 ;
   Valve[20].ZSOverride := 1 ;
   Valve[20].Ports := 0 ;
   Valve[20].PriorityCfg := 0 ;
   Valve[20].ZSOpenEnable := 0 ;
   Valve[20].Alarm := 0 ;
   Valve[20].ZSCloseEnable := 0 ;
   Valve[20].ZSOpenAddress := 0 ;
   Valve[20].ZSCloseAddress := 0 ;
   Valve[20].OutputAddress := 52 ;
   
   (*Reset Loop : Set to 0 the Valve[21 to 99].EnableCfg
   ============================================================*)
   FOR Config.IndeXValve := 21 to 99 by 1 do
   	Valve[Config.IndeXValve].EnableCfg := 0 ;
   	Valve[Config.IndeXValve].Alarm := 0 ;
   	Valve[Config.IndeXValve].Control := 0 ;
   	Valve[Config.IndeXValve].Auto := 0 ;
   	Valve[Config.IndeXValve].Manual := 0 ;
   	Valve[Config.IndeXValve].StatusWord := 0 ;
   	Valve[Config.IndeXValve].Status := 0 ;
   End_for ;
END_ROUTINE

ROUTINE Control_Loop   (* ladder *)
// Control Loop Routine
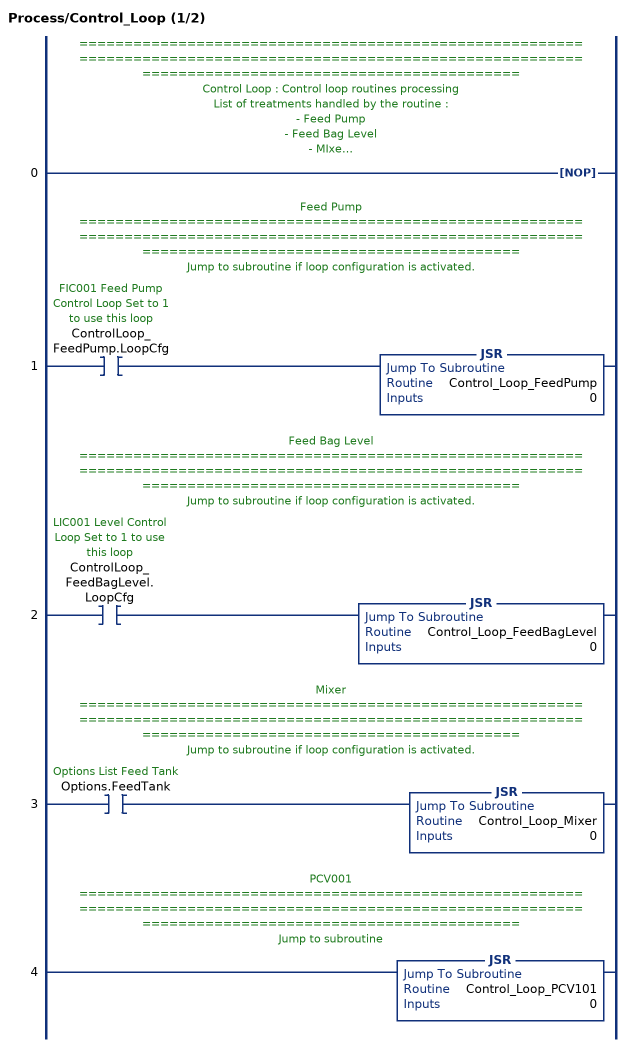
   // ==========================================================================================================================================================
   //                                                                                                                 Control Loop : Control loop routines processing
   //                                                     List of treatments handled by the routine :
   //                                                          - Feed Pump
   //                                                          - Feed Bag Level
   //                                                          - MIxer
   //                                                          - PCV001
   //                                                           - PCV101
   //                                                          - TIC101
   //                                                     -----------------------------------------------------------------------------------------------------------------------------------------------------
   //                                                     History
   // 		2019-DEC-24 - Merck - Q. Spindler - Initial version for Candidate Release 1.00.00.00.a
   // ==========================================================================================================================================================
   0: NOP();
   // Feed Pump
   // ==========================================================================================================================================================
   // Jump to subroutine if loop configuration is activated.
   1: XIC(ControlLoop_FeedPump.LoopCfg)JSR(Control_Loop_FeedPump,0);
   // Feed Bag Level
   // ==========================================================================================================================================================
   // Jump to subroutine if loop configuration is activated.
   2: XIC(ControlLoop_FeedBagLevel.LoopCfg)JSR(Control_Loop_FeedBagLevel,0);
   // Mixer
   // ==========================================================================================================================================================
   // Jump to subroutine if loop configuration is activated.
   3: XIC(Options.FeedTank)JSR(Control_Loop_Mixer,0);
   // PCV001
   // ==========================================================================================================================================================
   // Jump to subroutine
   4: JSR(Control_Loop_PCV101,0);
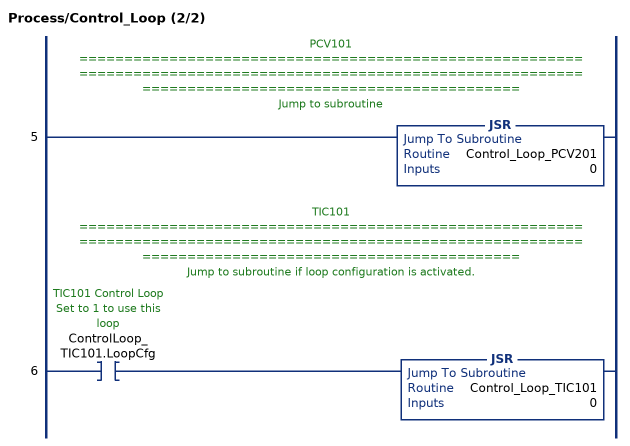
   // PCV101
   // ==========================================================================================================================================================
   // Jump to subroutine
   5: JSR(Control_Loop_PCV201,0);
   // TIC101
   // ==========================================================================================================================================================
   // Jump to subroutine if loop configuration is activated.
   6: XIC(ControlLoop_TIC101.LoopCfg)JSR(Control_Loop_TIC101,0);
END_ROUTINE

ROUTINE Control_Loop_FeedBagLevel   (* ladder *)
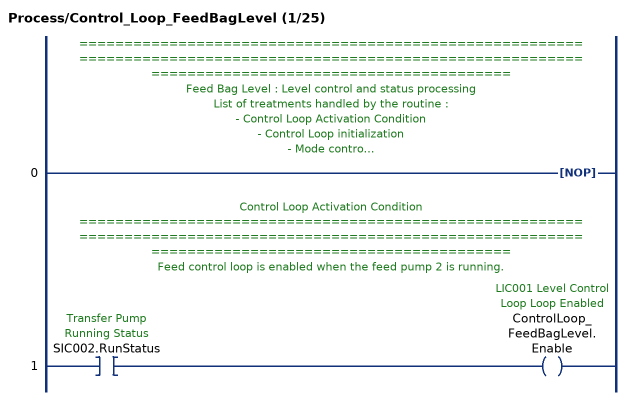
   // ========================================================================================================================================================
   //                                                                                                       Feed Bag Level : Level control and status processing
   //                                                     List of treatments handled by the routine :
   //                                                          - Control Loop Activation Condition
   //                                                          - Control Loop initialization
   //                                                          - Mode control
   //                                                          - Control Loop deadband calculation
   //                                                          - Management of ramping control
   //                                                          - Control Loop Stability control
   //                                                          - Control Loop manual state control
   //                                                          - Management of PID instruction
   //                                                          - Control of the analog output
   //                                                     -----------------------------------------------------------------------------------------------------------------------------------------------------
   //                                                     History
   //                		2019-DEC-24 - Merck - Q. Spindler - Initial version for Candidate Release 1.00.00.00.a
   // 		2020-SEP-09 - Merck - Q. Spindler - Modifications for Candidate Release 1.00.00.00.d
   // 					- Add ControlLoop Enable and not manual condition for DBOK status
   //                    - Set ramp rate minimum to 0.1
   // 		2021-APR-16 - Merck - Q. Spindler - Modifications for Candidate Release 1.00.00.00.e
   //                                        - Add Initialize address if no mode selected.
   //                                                              - The wrong control loop was used in the PID initialisation
   // 		2022-NOV-21 - Actemium - J. Jaekel - Modifications for Candidate Release 1.01.00.01.b
   // - Set manuel mode if Auto Mode 2 is enabled and TransferFlow option is disabled.
   // - If no mode is active, activate the manual mode.
   // ========================================================================================================================================================
   0: NOP();
   // Control Loop Activation Condition
   // ========================================================================================================================================================
   // Feed control loop is enabled when the feed pump 2 is running.
   1: XIC(SIC002.RunStatus)OTE(ControlLoop_FeedBagLevel.Enable);
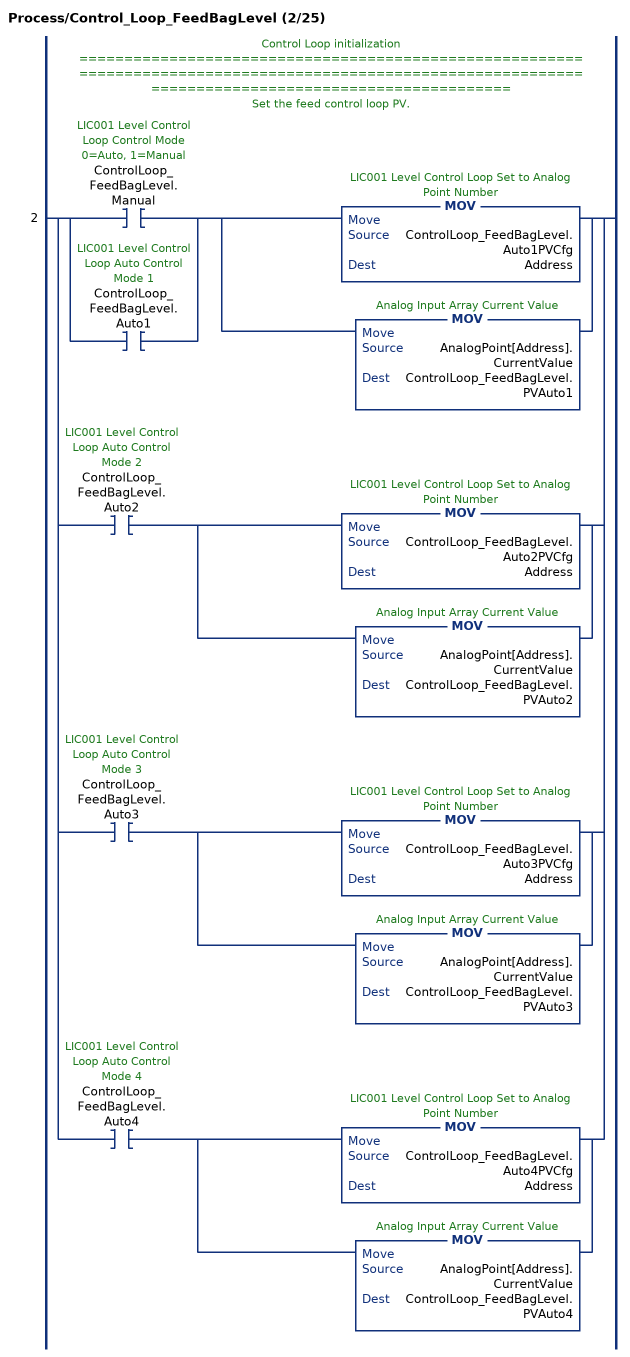
   // Control Loop initialization
   // ========================================================================================================================================================
   // Set the feed control loop PV.
   2: [[[XIC(ControlLoop_FeedBagLevel.Manual) ,XIC(ControlLoop_FeedBagLevel.Auto1) ] [MOV(ControlLoop_FeedBagLevel.Auto1PVCfg,Address) ,MOV(AnalogPoint[Address].CurrentValue,ControlLoop_FeedBagLevel.PVAuto1) ] ,XIC(ControlLoop_FeedBagLevel.Auto2) [MOV(ControlLoop_FeedBagLevel.Auto2PVCfg,Address) ,MOV(AnalogPoint[Address].CurrentValue,ControlLoop_FeedBagLevel.PVAuto2) ] ] ,XIC(ControlLoop_FeedBagLevel.Auto3) [MOV(ControlLoop_FeedBagLevel.Auto3PVCfg,Address) ,MOV(AnalogPoint[Address].CurrentValue,ControlLoop_FeedBagLevel.PVAuto3) ] ,XIC(ControlLoop_FeedBagLevel.Auto4) [MOV(ControlLoop_FeedBagLevel.Auto4PVCfg,Address) ,MOV(AnalogPoint[Address].CurrentValue,ControlLoop_FeedBagLevel.PVAuto4) ] ];
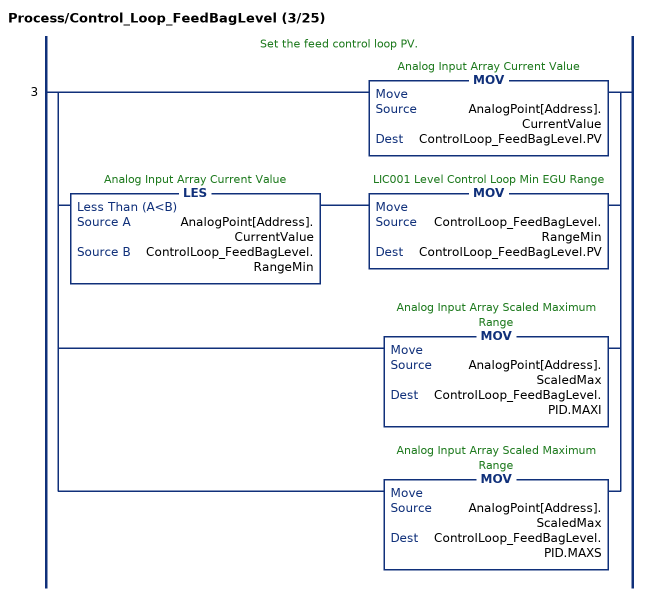
   // Set the feed control loop PV.
   3: [MOV(AnalogPoint[Address].CurrentValue,ControlLoop_FeedBagLevel.PV) ,LES(AnalogPoint[Address].CurrentValue,ControlLoop_FeedBagLevel.RangeMin) MOV(ControlLoop_FeedBagLevel.RangeMin,ControlLoop_FeedBagLevel.PV) ,MOV(AnalogPoint[Address].ScaledMax,ControlLoop_FeedBagLevel.PID.MAXI) ,MOV(AnalogPoint[Address].ScaledMax,ControlLoop_FeedBagLevel.PID.MAXS) ];
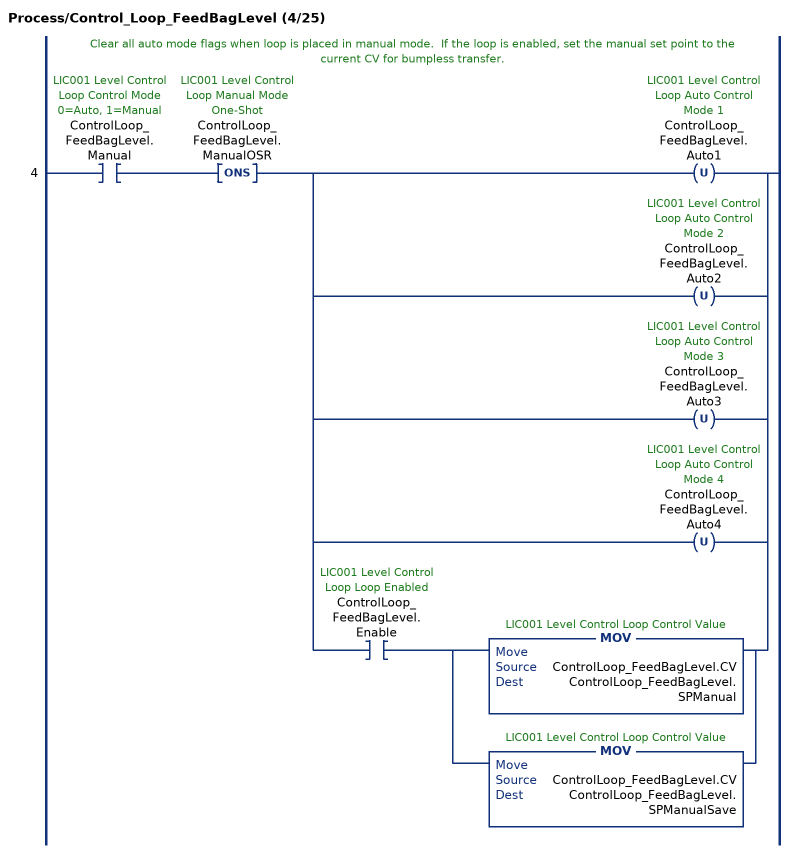
   // Clear all auto mode flags when loop is placed in manual mode.  If the loop is enabled, set the manual set point to the current CV for bumpless transfer.
   4: XIC(ControlLoop_FeedBagLevel.Manual)ONS(ControlLoop_FeedBagLevel.ManualOSR)[OTU(ControlLoop_FeedBagLevel.Auto1) ,OTU(ControlLoop_FeedBagLevel.Auto2) ,OTU(ControlLoop_FeedBagLevel.Auto3) ,OTU(ControlLoop_FeedBagLevel.Auto4) ,XIC(ControlLoop_FeedBagLevel.Enable) [MOV(ControlLoop_FeedBagLevel.CV,ControlLoop_FeedBagLevel.SPManual) ,MOV(ControlLoop_FeedBagLevel.CV,ControlLoop_FeedBagLevel.SPManualSave) ] ];
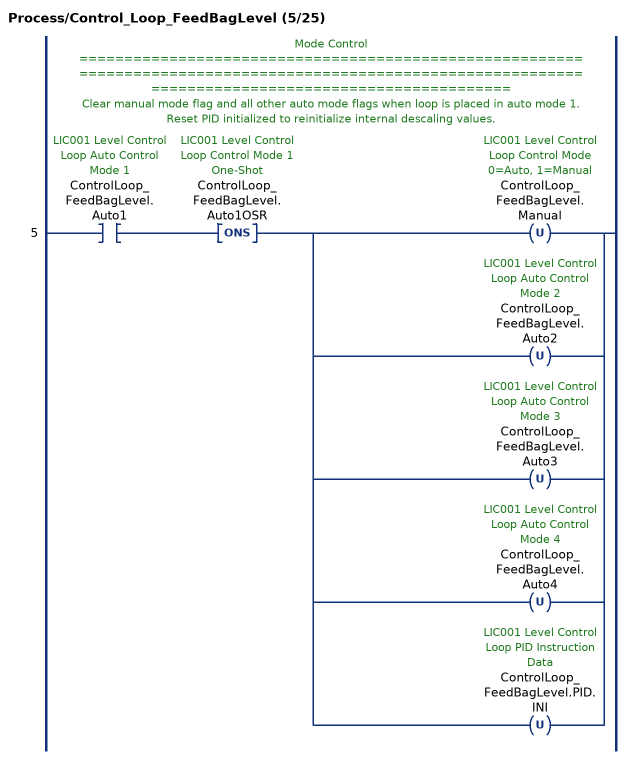
   // Mode Control
   // ========================================================================================================================================================
   // Clear manual mode flag and all other auto mode flags when loop is placed in auto mode 1. Reset PID initialized to reinitialize internal descaling values.
   5: XIC(ControlLoop_FeedBagLevel.Auto1)ONS(ControlLoop_FeedBagLevel.Auto1OSR)[OTU(ControlLoop_FeedBagLevel.Manual) ,OTU(ControlLoop_FeedBagLevel.Auto2) ,OTU(ControlLoop_FeedBagLevel.Auto3) ,OTU(ControlLoop_FeedBagLevel.Auto4) ,OTU(ControlLoop_FeedBagLevel.PID.INI) ];
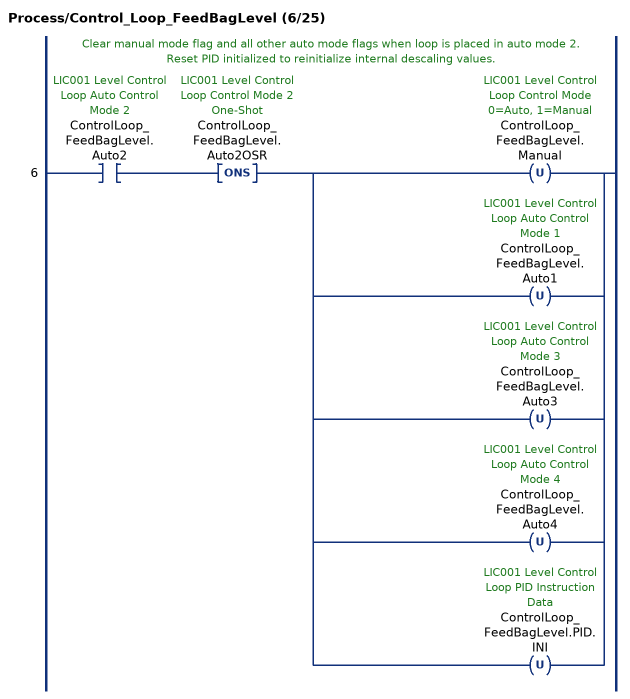
   // Clear manual mode flag and all other auto mode flags when loop is placed in auto mode 2. Reset PID initialized to reinitialize internal descaling values.
   6: XIC(ControlLoop_FeedBagLevel.Auto2)ONS(ControlLoop_FeedBagLevel.Auto2OSR)[OTU(ControlLoop_FeedBagLevel.Manual) ,OTU(ControlLoop_FeedBagLevel.Auto1) ,OTU(ControlLoop_FeedBagLevel.Auto3) ,OTU(ControlLoop_FeedBagLevel.Auto4) ,OTU(ControlLoop_FeedBagLevel.PID.INI) ];
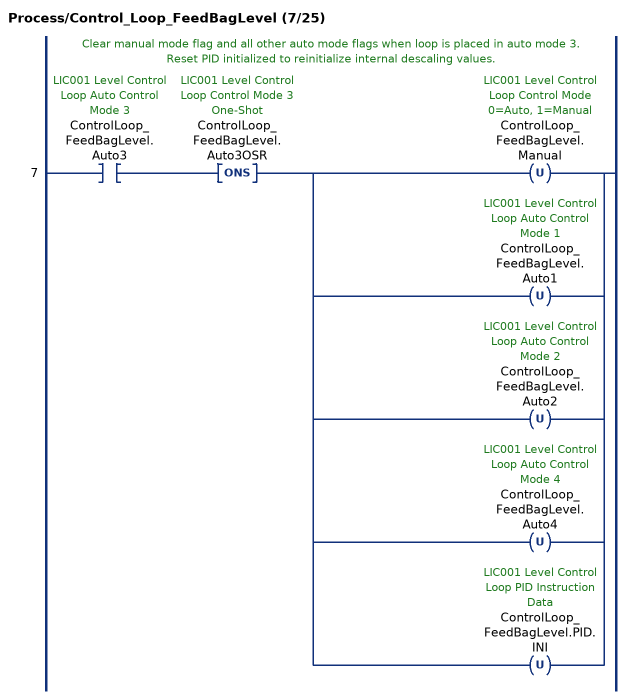
   // Clear manual mode flag and all other auto mode flags when loop is placed in auto mode 3. Reset PID initialized to reinitialize internal descaling values.
   7: XIC(ControlLoop_FeedBagLevel.Auto3)ONS(ControlLoop_FeedBagLevel.Auto3OSR)[OTU(ControlLoop_FeedBagLevel.Manual) ,OTU(ControlLoop_FeedBagLevel.Auto1) ,OTU(ControlLoop_FeedBagLevel.Auto2) ,OTU(ControlLoop_FeedBagLevel.Auto4) ,OTU(ControlLoop_FeedBagLevel.PID.INI) ];
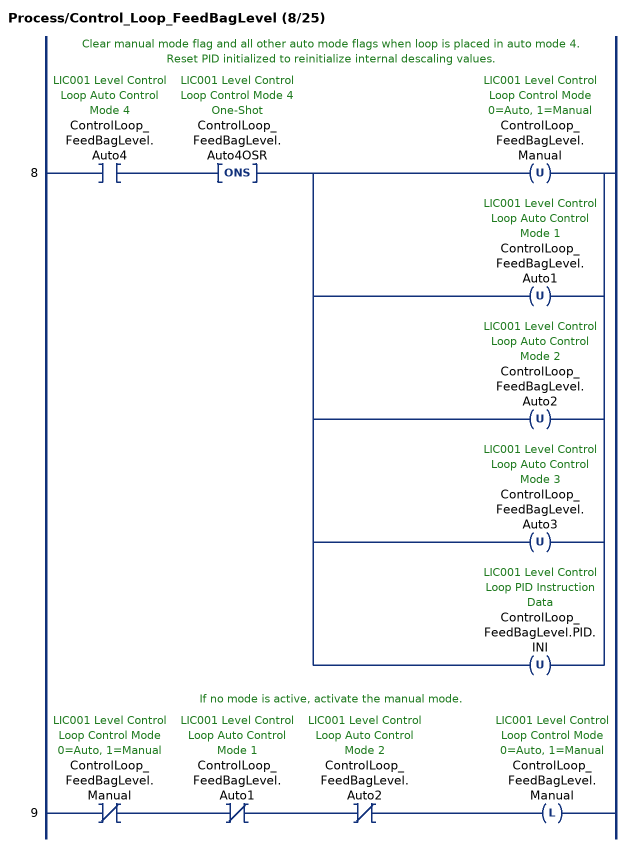
   // Clear manual mode flag and all other auto mode flags when loop is placed in auto mode 4. Reset PID initialized to reinitialize internal descaling values.
   8: XIC(ControlLoop_FeedBagLevel.Auto4)ONS(ControlLoop_FeedBagLevel.Auto4OSR)[OTU(ControlLoop_FeedBagLevel.Manual) ,OTU(ControlLoop_FeedBagLevel.Auto1) ,OTU(ControlLoop_FeedBagLevel.Auto2) ,OTU(ControlLoop_FeedBagLevel.Auto3) ,OTU(ControlLoop_FeedBagLevel.PID.INI) ];
   // If no mode is active, activate the manual mode.
   9: XIO(ControlLoop_FeedBagLevel.Manual)XIO(ControlLoop_FeedBagLevel.Auto1)XIO(ControlLoop_FeedBagLevel.Auto2)OTL(ControlLoop_FeedBagLevel.Manual);
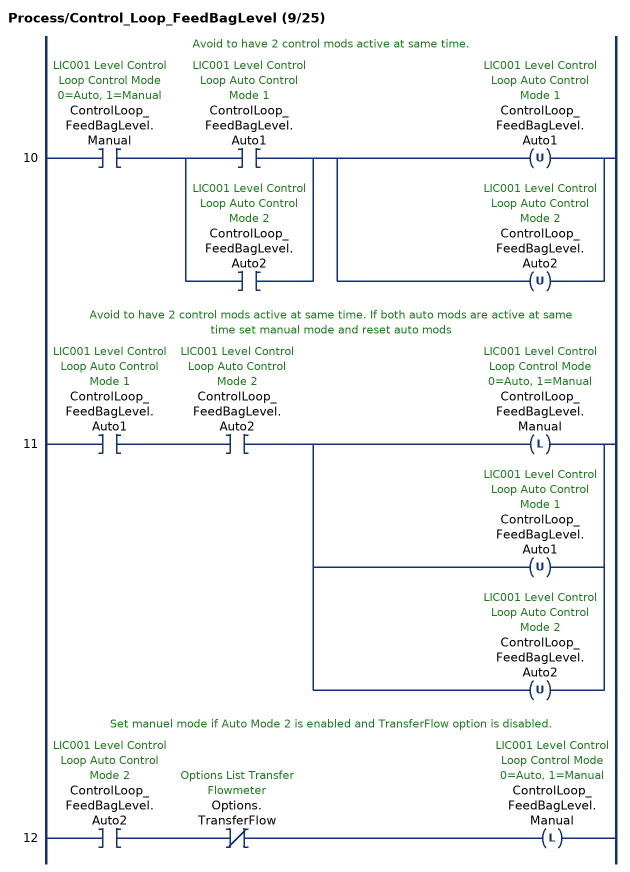
   // Avoid to have 2 control mods active at same time.
   10: XIC(ControlLoop_FeedBagLevel.Manual)[XIC(ControlLoop_FeedBagLevel.Auto1) ,XIC(ControlLoop_FeedBagLevel.Auto2) ][OTU(ControlLoop_FeedBagLevel.Auto1) ,OTU(ControlLoop_FeedBagLevel.Auto2) ];
   // Avoid to have 2 control mods active at same time. If both auto mods are active at same time set manual mode and reset auto mods
   11: XIC(ControlLoop_FeedBagLevel.Auto1)XIC(ControlLoop_FeedBagLevel.Auto2)[OTL(ControlLoop_FeedBagLevel.Manual) ,OTU(ControlLoop_FeedBagLevel.Auto1) ,OTU(ControlLoop_FeedBagLevel.Auto2) ];
   // Set manuel mode if Auto Mode 2 is enabled and TransferFlow option is disabled.
   12: XIC(ControlLoop_FeedBagLevel.Auto2)XIO(Options.TransferFlow)OTL(ControlLoop_FeedBagLevel.Manual);
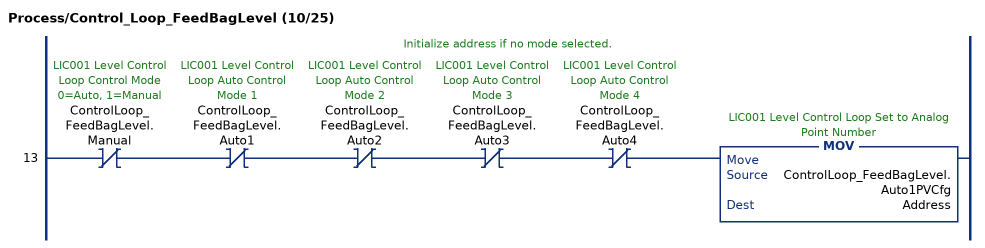
   // Initialize address if no mode selected.
   13: XIO(ControlLoop_FeedBagLevel.Manual)XIO(ControlLoop_FeedBagLevel.Auto1)XIO(ControlLoop_FeedBagLevel.Auto2)XIO(ControlLoop_FeedBagLevel.Auto3)XIO(ControlLoop_FeedBagLevel.Auto4)MOV(ControlLoop_FeedBagLevel.Auto1PVCfg,Address);
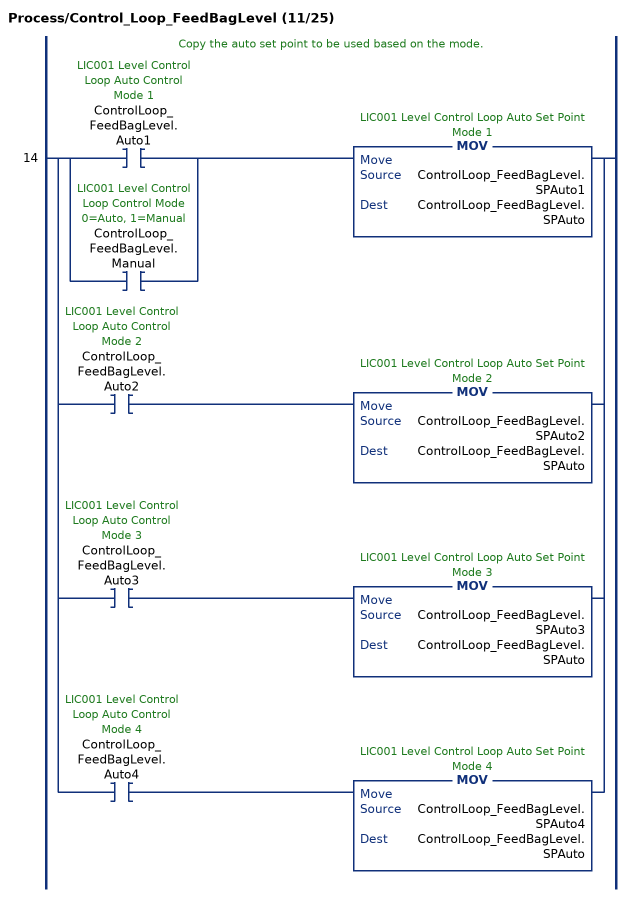
   // Copy the auto set point to be used based on the mode.
   14: [[XIC(ControlLoop_FeedBagLevel.Auto1) ,XIC(ControlLoop_FeedBagLevel.Manual) ] MOV(ControlLoop_FeedBagLevel.SPAuto1,ControlLoop_FeedBagLevel.SPAuto) ,XIC(ControlLoop_FeedBagLevel.Auto2) MOV(ControlLoop_FeedBagLevel.SPAuto2,ControlLoop_FeedBagLevel.SPAuto) ,XIC(ControlLoop_FeedBagLevel.Auto3) MOV(ControlLoop_FeedBagLevel.SPAuto3,ControlLoop_FeedBagLevel.SPAuto) ,XIC(ControlLoop_FeedBagLevel.Auto4) MOV(ControlLoop_FeedBagLevel.SPAuto4,ControlLoop_FeedBagLevel.SPAuto) ];
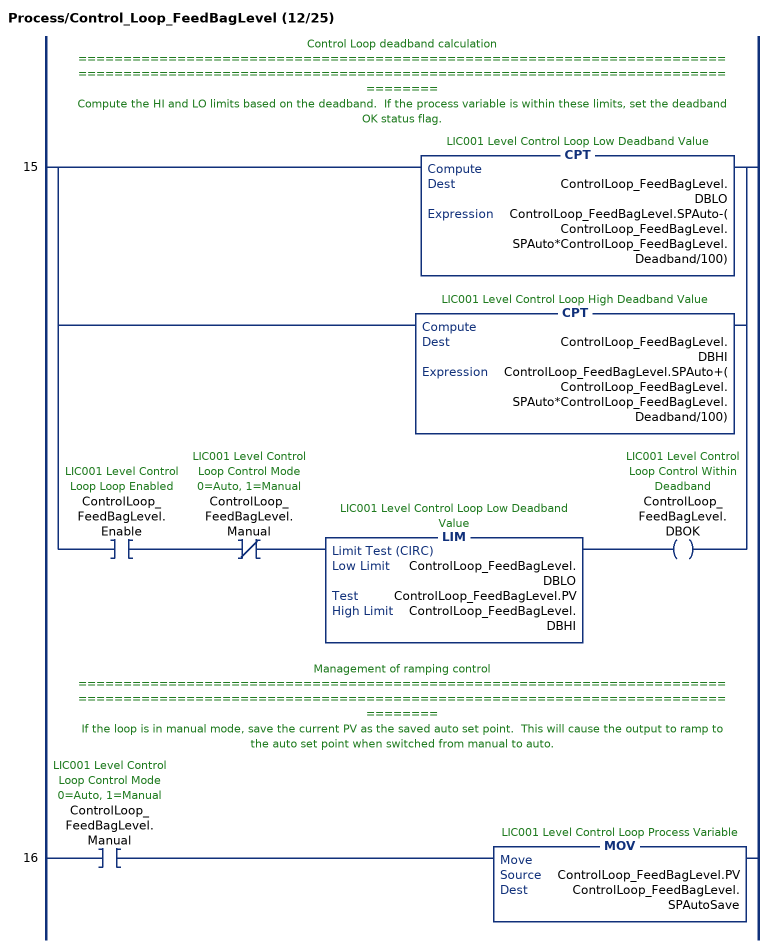
   // Control Loop deadband calculation
   // ========================================================================================================================================================
   // Compute the HI and LO limits based on the deadband.  If the process variable is within these limits, set the deadband OK status flag.
   15: [CPT(ControlLoop_FeedBagLevel.DBLO,ControlLoop_FeedBagLevel.SPAuto-(ControlLoop_FeedBagLevel.SPAuto*ControlLoop_FeedBagLevel.Deadband/100)) ,CPT(ControlLoop_FeedBagLevel.DBHI,ControlLoop_FeedBagLevel.SPAuto+(ControlLoop_FeedBagLevel.SPAuto*ControlLoop_FeedBagLevel.Deadband/100)) ,XIC(ControlLoop_FeedBagLevel.Enable) XIO(ControlLoop_FeedBagLevel.Manual) LIM(ControlLoop_FeedBagLevel.DBLO,ControlLoop_FeedBagLevel.PV,ControlLoop_FeedBagLevel.DBHI) OTE(ControlLoop_FeedBagLevel.DBOK) ];
   // Management of ramping control
   // ========================================================================================================================================================
   // If the loop is in manual mode, save the current PV as the saved auto set point.  This will cause the output to ramp to the auto set point when switched from manual to auto.
   16: XIC(ControlLoop_FeedBagLevel.Manual)MOV(ControlLoop_FeedBagLevel.PV,ControlLoop_FeedBagLevel.SPAutoSave);
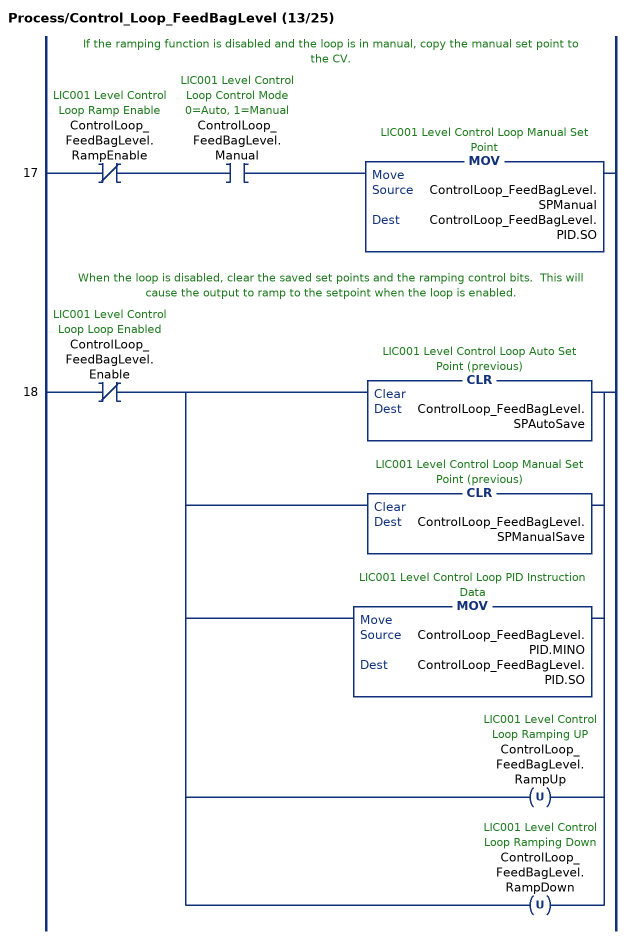
   // If the ramping function is disabled and the loop is in manual, copy the manual set point to the CV.
   17: XIO(ControlLoop_FeedBagLevel.RampEnable)XIC(ControlLoop_FeedBagLevel.Manual)MOV(ControlLoop_FeedBagLevel.SPManual,ControlLoop_FeedBagLevel.PID.SO);
   // When the loop is disabled, clear the saved set points and the ramping control bits.  This will cause the output to ramp to the setpoint when the loop is enabled.
   18: XIO(ControlLoop_FeedBagLevel.Enable)[CLR(ControlLoop_FeedBagLevel.SPAutoSave) ,CLR(ControlLoop_FeedBagLevel.SPManualSave) ,MOV(ControlLoop_FeedBagLevel.PID.MINO,ControlLoop_FeedBagLevel.PID.SO) ,OTU(ControlLoop_FeedBagLevel.RampUp) ,OTU(ControlLoop_FeedBagLevel.RampDown) ];
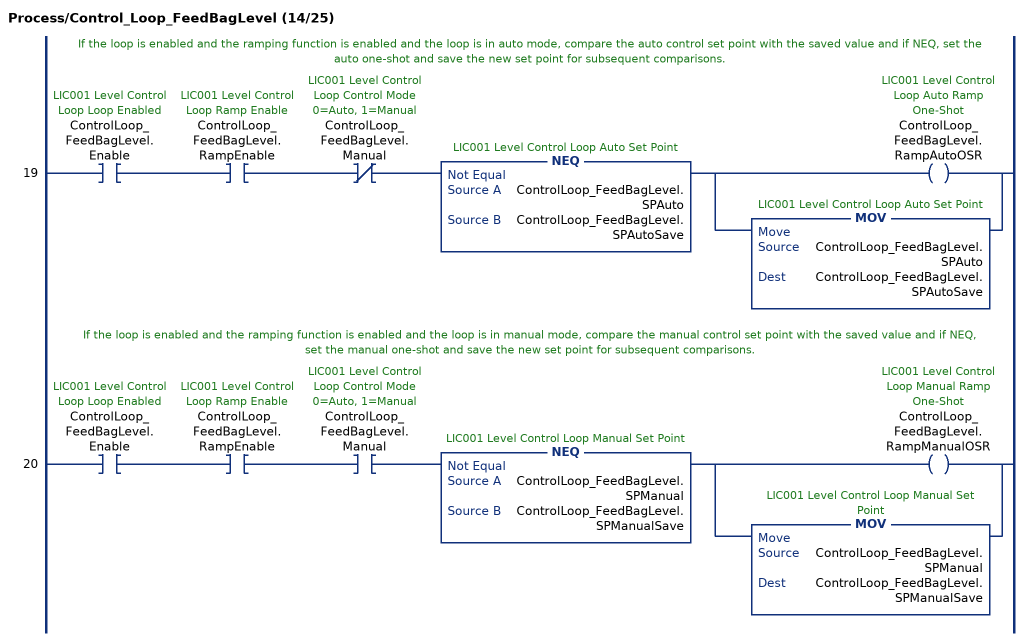
   // If the loop is enabled and the ramping function is enabled and the loop is in auto mode, compare the auto control set point with the saved value and if NEQ, set the auto one-shot and save the new set point for subsequent comparisons.
   19: XIC(ControlLoop_FeedBagLevel.Enable)XIC(ControlLoop_FeedBagLevel.RampEnable)XIO(ControlLoop_FeedBagLevel.Manual)NEQ(ControlLoop_FeedBagLevel.SPAuto,ControlLoop_FeedBagLevel.SPAutoSave)[OTE(ControlLoop_FeedBagLevel.RampAutoOSR) ,MOV(ControlLoop_FeedBagLevel.SPAuto,ControlLoop_FeedBagLevel.SPAutoSave) ];
   // If the loop is enabled and the ramping function is enabled and the loop is in manual mode, compare the manual control set point with the saved value and if NEQ, set the manual one-shot and save the new set point for subsequent comparisons.
   20: XIC(ControlLoop_FeedBagLevel.Enable)XIC(ControlLoop_FeedBagLevel.RampEnable)XIC(ControlLoop_FeedBagLevel.Manual)NEQ(ControlLoop_FeedBagLevel.SPManual,ControlLoop_FeedBagLevel.SPManualSave)[OTE(ControlLoop_FeedBagLevel.RampManualOSR) ,MOV(ControlLoop_FeedBagLevel.SPManual,ControlLoop_FeedBagLevel.SPManualSave) ];
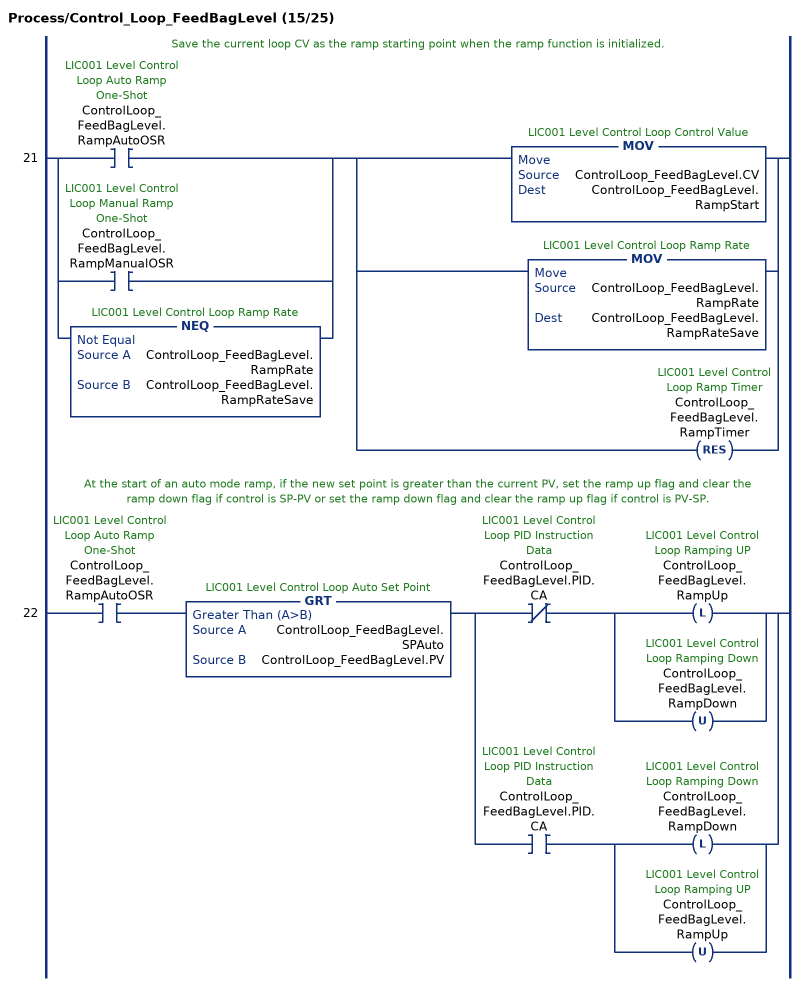
   // Save the current loop CV as the ramp starting point when the ramp function is initialized.
   21: [XIC(ControlLoop_FeedBagLevel.RampAutoOSR) ,XIC(ControlLoop_FeedBagLevel.RampManualOSR) ,NEQ(ControlLoop_FeedBagLevel.RampRate,ControlLoop_FeedBagLevel.RampRateSave) ][MOV(ControlLoop_FeedBagLevel.CV,ControlLoop_FeedBagLevel.RampStart) ,MOV(ControlLoop_FeedBagLevel.RampRate,ControlLoop_FeedBagLevel.RampRateSave) ,RES(ControlLoop_FeedBagLevel.RampTimer) ];
   // At the start of an auto mode ramp, if the new set point is greater than the current PV, set the ramp up flag and clear the ramp down flag if control is SP-PV or set the ramp down flag and clear the ramp up flag if control is PV-SP.
   22: XIC(ControlLoop_FeedBagLevel.RampAutoOSR)GRT(ControlLoop_FeedBagLevel.SPAuto,ControlLoop_FeedBagLevel.PV)[XIO(ControlLoop_FeedBagLevel.PID.CA) [OTL(ControlLoop_FeedBagLevel.RampUp) ,OTU(ControlLoop_FeedBagLevel.RampDown) ] ,XIC(ControlLoop_FeedBagLevel.PID.CA) [OTL(ControlLoop_FeedBagLevel.RampDown) ,OTU(ControlLoop_FeedBagLevel.RampUp) ] ];
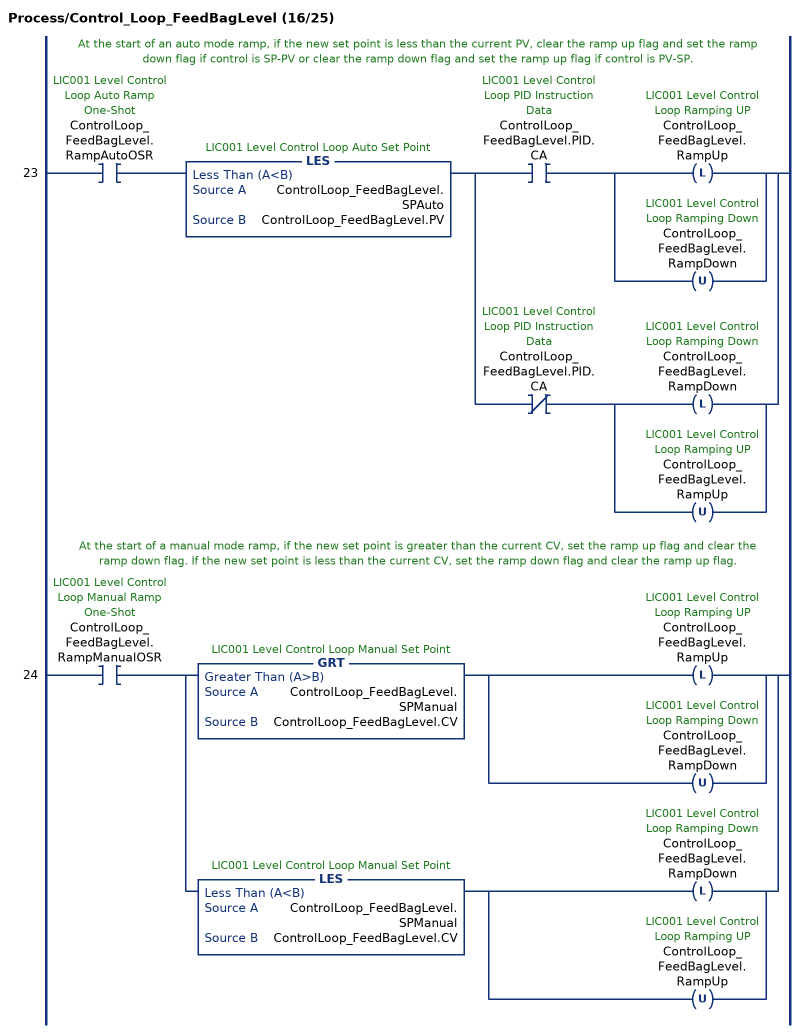
   // At the start of an auto mode ramp, if the new set point is less than the current PV, clear the ramp up flag and set the ramp down flag if control is SP-PV or clear the ramp down flag and set the ramp up flag if control is PV-SP.
   23: XIC(ControlLoop_FeedBagLevel.RampAutoOSR)LES(ControlLoop_FeedBagLevel.SPAuto,ControlLoop_FeedBagLevel.PV)[XIC(ControlLoop_FeedBagLevel.PID.CA) [OTL(ControlLoop_FeedBagLevel.RampUp) ,OTU(ControlLoop_FeedBagLevel.RampDown) ] ,XIO(ControlLoop_FeedBagLevel.PID.CA) [OTL(ControlLoop_FeedBagLevel.RampDown) ,OTU(ControlLoop_FeedBagLevel.RampUp) ] ];
   // At the start of a manual mode ramp, if the new set point is greater than the current CV, set the ramp up flag and clear the ramp down flag. If the new set point is less than the current CV, set the ramp down flag and clear the ramp up flag.
   24: XIC(ControlLoop_FeedBagLevel.RampManualOSR)[GRT(ControlLoop_FeedBagLevel.SPManual,ControlLoop_FeedBagLevel.CV) [OTL(ControlLoop_FeedBagLevel.RampUp) ,OTU(ControlLoop_FeedBagLevel.RampDown) ] ,LES(ControlLoop_FeedBagLevel.SPManual,ControlLoop_FeedBagLevel.CV) [OTL(ControlLoop_FeedBagLevel.RampDown) ,OTU(ControlLoop_FeedBagLevel.RampUp) ] ];
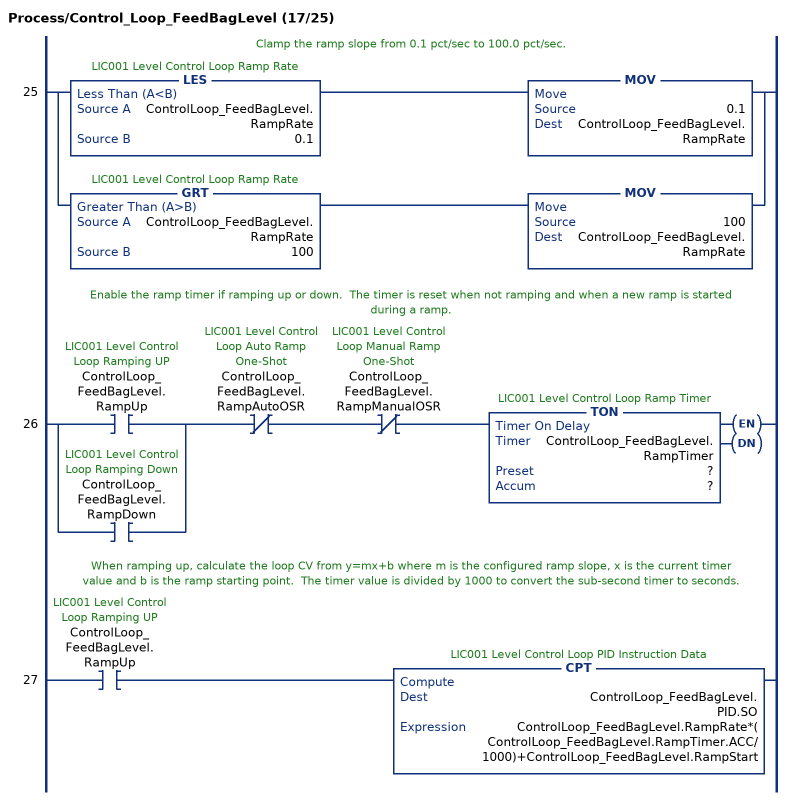
   // Clamp the ramp slope from 0.1 pct/sec to 100.0 pct/sec.
   25: [LES(ControlLoop_FeedBagLevel.RampRate,0.1) MOV(0.1,ControlLoop_FeedBagLevel.RampRate) ,GRT(ControlLoop_FeedBagLevel.RampRate,100) MOV(100,ControlLoop_FeedBagLevel.RampRate) ];
   // Enable the ramp timer if ramping up or down.  The timer is reset when not ramping and when a new ramp is started during a ramp.
   26: [XIC(ControlLoop_FeedBagLevel.RampUp) ,XIC(ControlLoop_FeedBagLevel.RampDown) ]XIO(ControlLoop_FeedBagLevel.RampAutoOSR)XIO(ControlLoop_FeedBagLevel.RampManualOSR)TON(ControlLoop_FeedBagLevel.RampTimer,?,?);
   // When ramping up, calculate the loop CV from y=mx+b where m is the configured ramp slope, x is the current timer value and b is the ramp starting point.  The timer value is divided by 1000 to convert the sub-second timer to seconds.
   27: XIC(ControlLoop_FeedBagLevel.RampUp)CPT(ControlLoop_FeedBagLevel.PID.SO,ControlLoop_FeedBagLevel.RampRate*(ControlLoop_FeedBagLevel.RampTimer.ACC/1000)+ControlLoop_FeedBagLevel.RampStart);
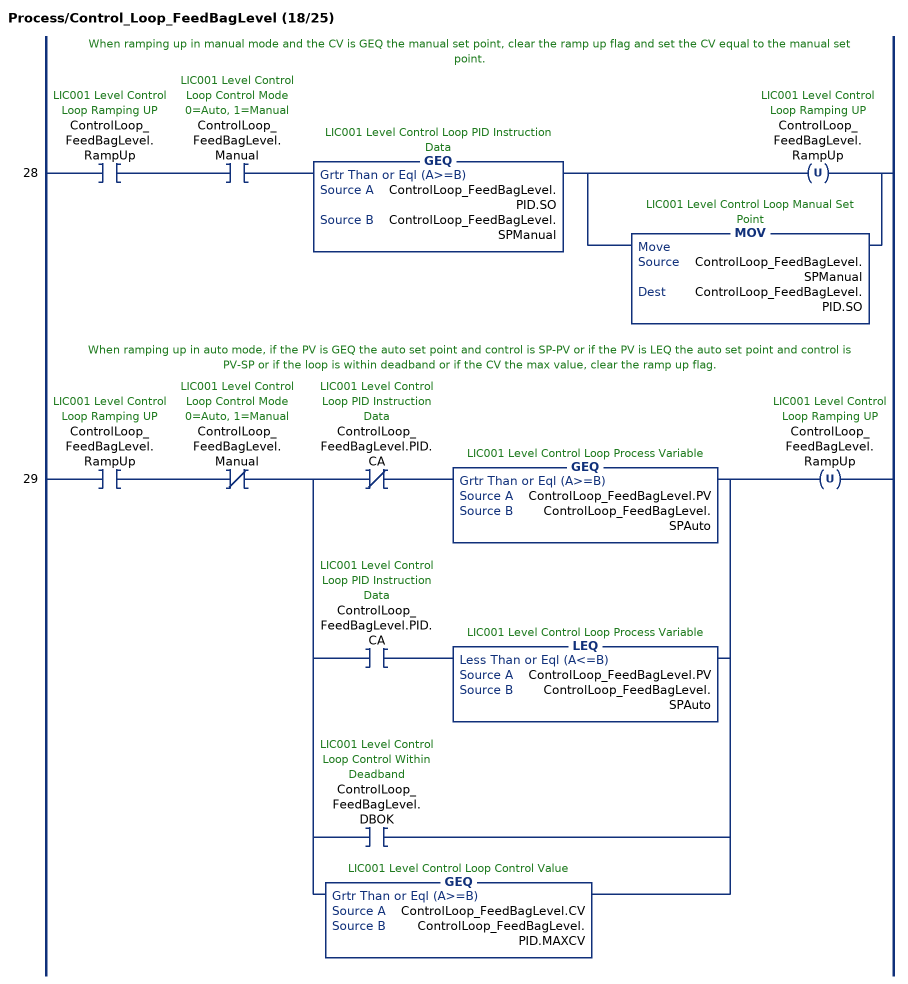
   // When ramping up in manual mode and the CV is GEQ the manual set point, clear the ramp up flag and set the CV equal to the manual set point.
   28: XIC(ControlLoop_FeedBagLevel.RampUp)XIC(ControlLoop_FeedBagLevel.Manual)GEQ(ControlLoop_FeedBagLevel.PID.SO,ControlLoop_FeedBagLevel.SPManual)[OTU(ControlLoop_FeedBagLevel.RampUp) ,MOV(ControlLoop_FeedBagLevel.SPManual,ControlLoop_FeedBagLevel.PID.SO) ];
   // When ramping up in auto mode, if the PV is GEQ the auto set point and control is SP-PV or if the PV is LEQ the auto set point and control is PV-SP or if the loop is within deadband or if the CV the max value, clear the ramp up flag.
   29: XIC(ControlLoop_FeedBagLevel.RampUp)XIO(ControlLoop_FeedBagLevel.Manual)[XIO(ControlLoop_FeedBagLevel.PID.CA) GEQ(ControlLoop_FeedBagLevel.PV,ControlLoop_FeedBagLevel.SPAuto) ,XIC(ControlLoop_FeedBagLevel.PID.CA) LEQ(ControlLoop_FeedBagLevel.PV,ControlLoop_FeedBagLevel.SPAuto) ,XIC(ControlLoop_FeedBagLevel.DBOK) ,GEQ(ControlLoop_FeedBagLevel.CV,ControlLoop_FeedBagLevel.PID.MAXCV) ]OTU(ControlLoop_FeedBagLevel.RampUp);
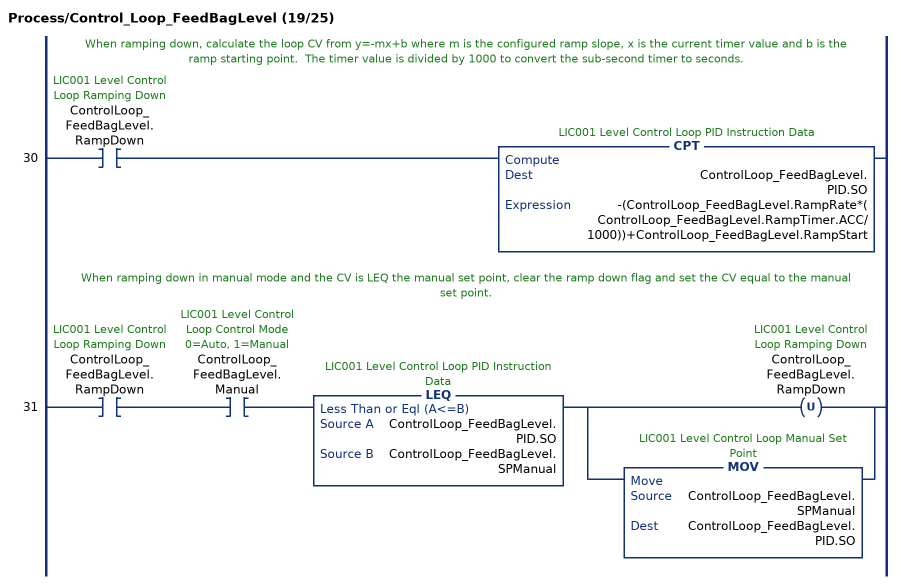
   // When ramping down, calculate the loop CV from y=-mx+b where m is the configured ramp slope, x is the current timer value and b is the ramp starting point.  The timer value is divided by 1000 to convert the sub-second timer to seconds.
   30: XIC(ControlLoop_FeedBagLevel.RampDown)CPT(ControlLoop_FeedBagLevel.PID.SO,-(ControlLoop_FeedBagLevel.RampRate*(ControlLoop_FeedBagLevel.RampTimer.ACC/1000))+ControlLoop_FeedBagLevel.RampStart);
   // When ramping down in manual mode and the CV is LEQ the manual set point, clear the ramp down flag and set the CV equal to the manual set point.
   31: XIC(ControlLoop_FeedBagLevel.RampDown)XIC(ControlLoop_FeedBagLevel.Manual)LEQ(ControlLoop_FeedBagLevel.PID.SO,ControlLoop_FeedBagLevel.SPManual)[OTU(ControlLoop_FeedBagLevel.RampDown) ,MOV(ControlLoop_FeedBagLevel.SPManual,ControlLoop_FeedBagLevel.PID.SO) ];
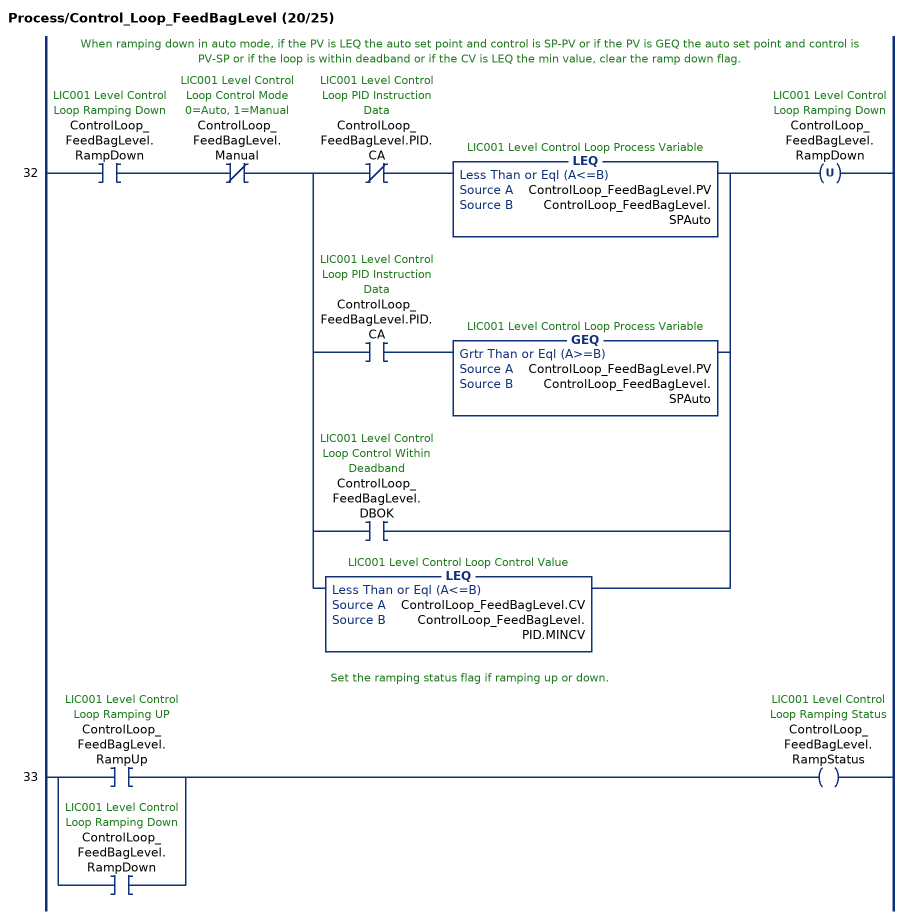
   // When ramping down in auto mode, if the PV is LEQ the auto set point and control is SP-PV or if the PV is GEQ the auto set point and control is PV-SP or if the loop is within deadband or if the CV is LEQ the min value, clear the ramp down flag.
   32: XIC(ControlLoop_FeedBagLevel.RampDown)XIO(ControlLoop_FeedBagLevel.Manual)[XIO(ControlLoop_FeedBagLevel.PID.CA) LEQ(ControlLoop_FeedBagLevel.PV,ControlLoop_FeedBagLevel.SPAuto) ,XIC(ControlLoop_FeedBagLevel.PID.CA) GEQ(ControlLoop_FeedBagLevel.PV,ControlLoop_FeedBagLevel.SPAuto) ,XIC(ControlLoop_FeedBagLevel.DBOK) ,LEQ(ControlLoop_FeedBagLevel.CV,ControlLoop_FeedBagLevel.PID.MINCV) ]OTU(ControlLoop_FeedBagLevel.RampDown);
   // Set the ramping status flag if ramping up or down.
   33: [XIC(ControlLoop_FeedBagLevel.RampUp) ,XIC(ControlLoop_FeedBagLevel.RampDown) ]OTE(ControlLoop_FeedBagLevel.RampStatus);
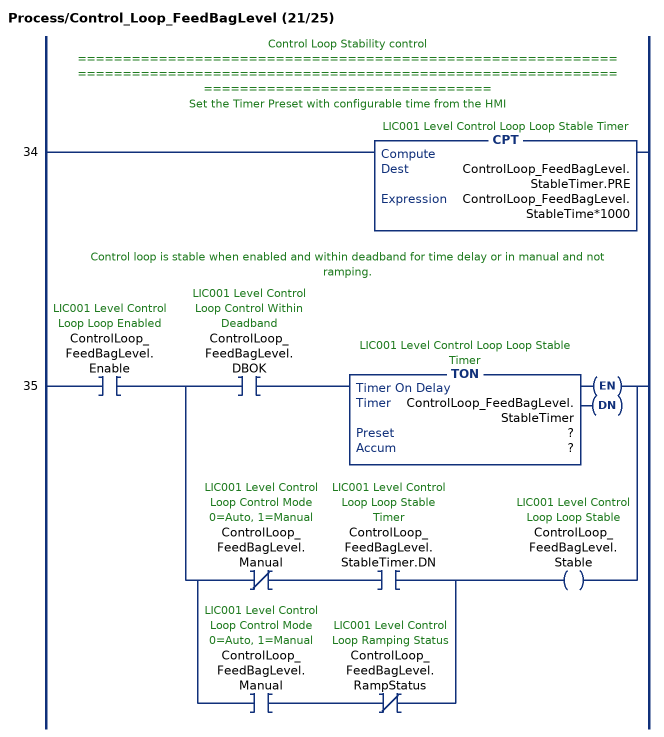
   // Control Loop Stability control
   // ========================================================================================================================================================
   // Set the Timer Preset with configurable time from the HMI
   34: CPT(ControlLoop_FeedBagLevel.StableTimer.PRE,ControlLoop_FeedBagLevel.StableTime*1000);
   // Control loop is stable when enabled and within deadband for time delay or in manual and not ramping.
   35: XIC(ControlLoop_FeedBagLevel.Enable)[XIC(ControlLoop_FeedBagLevel.DBOK) TON(ControlLoop_FeedBagLevel.StableTimer,?,?) ,[XIO(ControlLoop_FeedBagLevel.Manual) XIC(ControlLoop_FeedBagLevel.StableTimer.DN) ,XIC(ControlLoop_FeedBagLevel.Manual) XIO(ControlLoop_FeedBagLevel.RampStatus) ] OTE(ControlLoop_FeedBagLevel.Stable) ];
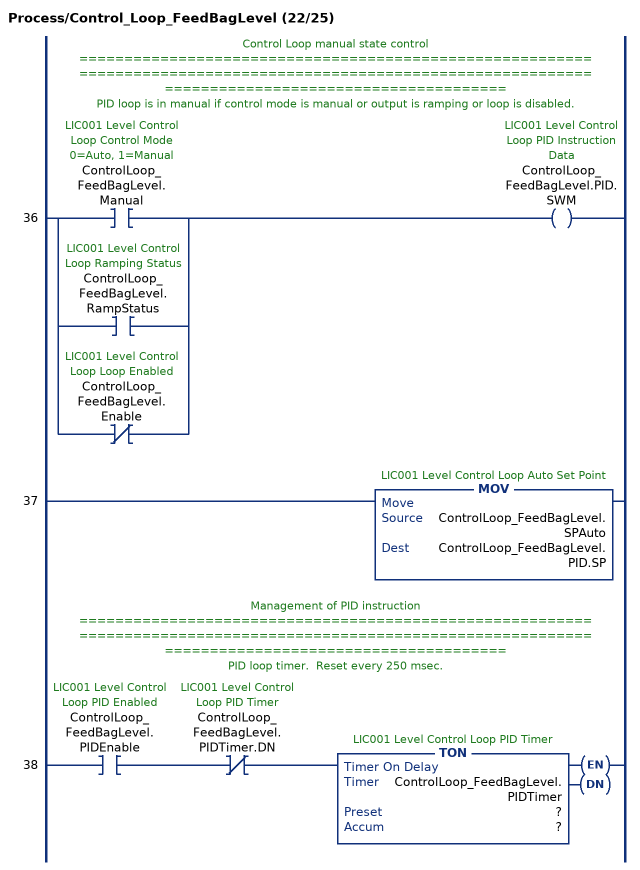
   // Control Loop manual state control
   // ========================================================================================================================================================
   // PID loop is in manual if control mode is manual or output is ramping or loop is disabled.
   36: [XIC(ControlLoop_FeedBagLevel.Manual) ,XIC(ControlLoop_FeedBagLevel.RampStatus) ,XIO(ControlLoop_FeedBagLevel.Enable) ]OTE(ControlLoop_FeedBagLevel.PID.SWM);
   37: MOV(ControlLoop_FeedBagLevel.SPAuto,ControlLoop_FeedBagLevel.PID.SP);
   // Management of PID instruction
   // ========================================================================================================================================================
   // PID loop timer.  Reset every 250 msec.
   38: XIC(ControlLoop_FeedBagLevel.PIDEnable)XIO(ControlLoop_FeedBagLevel.PIDTimer.DN)TON(ControlLoop_FeedBagLevel.PIDTimer,?,?);
